// TwinCAT 3 PLC project Syn_Visu_Demo
// ProgramVersion: 3.1.4026.28
// libraries:
//   SynConfig,2.4.0.0,Syntegon Group
//   SynVisu,10.0.0.0,Syntegon Group
//   Tc3_Module,newest,Beckhoff Automation GmbH
//   Tc2_System, * (Beckhoff Automation GmbH)
// project tree:
//   / DEMO_GlobalConst.TcGVL, DEMO_GlobalVar.TcGVL, GVL_Config.TcGVL, GVL_Visu.TcGVL, TVisuDemo_Detection.TcDUT, TVisuDemo_Recipe.TcDUT
//   POUs/ PlcTask.TcTTO, P_VisuDemo.TcPOU, P_VisuDemoCartesian.TcPOU, P_VisuDemoCartesianAxes.TcPOU, P_VisuDemoDelta.TcPOU, P_VisuDemoFxx.TcPOU, P_VisuDemoIdh.TcPOU, P_VisuDemoMachine.TcPOU, P_VisuDemoSpacing.TcPOU, P_VisuDemoStress.TcPOU, _FC_DemoApproach.TcPOU
// (motion and I/O tree: see PLC project syn_visu)
// real-time tasks:
//   TASK PlcTask: cycle T#10ms, priority 20, ADS port 350
//   TASK TestTask: cycle T#10ms, priority 21, ADS port 351

CONFIGURATION Syn_Visu_Demo
    RESOURCE PLC ON TwinCAT3
        TASK PlcTask(INTERVAL := T#10ms, PRIORITY := 20);
        PROGRAM P_VisuDemo WITH PlcTask : P_VisuDemo;
    END_RESOURCE
END_CONFIGURATION

// ---- TVisuDemo_Detection.TcDUT
(* A raw detection as the demo's product generator makes it up and a vision system would report it: where the
   product lies (MCS), the belt position at that moment and its type. The demo's tracking latches it as Vision 1's. *)
TYPE TVisuDemo_Detection :
STRUCT
	Pose								: ST_VisuPlanarPose;	// MCS
	lr_BeltPosition						: LREAL;	// [mm] Infeed 1's belt position when it was seen
	udn_ProductType						: UDINT;	// [-]
END_STRUCT
END_TYPE

// ---- TVisuDemo_Recipe.TcDUT
(* The demo's effective recipe (ADR 0022): what P_VisuDemoMachine reads from its Syn_Config machine FB every cycle
   and the Delta application runs with: Infeed 1's belt, Delta 1 and the product generator before Vision 1. *)
TYPE TVisuDemo_Recipe :
STRUCT
	lr_BeltSpeed						: LREAL;	// [mm/s] Infeed 1
	lr_BeltAccel						: LREAL;	// [mm/s2] Infeed 1, also its deceleration
	lr_RobotSpeed						: LREAL;	// [%] Delta 1, of its maximum TCP speed
	lr_RobotAccel						: LREAL;	// [%] Delta 1, of its maximum TCP acceleration
	dn_PicksPerCycle					: DINT;	// [-] Delta 1 picks this many products before it places them: 1 or 2
	lr_Rate								: LREAL;	// [1/min] places the generator fills per minute at the recipe's belt speed
	dn_Lanes							: DINT;	// [-] pattern Lanes: lanes across the belt, 1..4; each product goes into one at random
	lr_LanePitch						: LREAL;	// [mm] between the lanes, centred on the belt
	dn_TypeMix							: DINT;	// [-] 0 = every type, 1 = boxes, 2 = round (can, oval)
	lr_ScatterX							: LREAL;	// [mm] at most along the belt, either way
	lr_ScatterY							: LREAL;	// [mm] at most across the belt, either way
	lr_ScatterRz						: LREAL;	// [deg] at most turned, either way
	lr_GapShare							: LREAL;	// [%] of the generator's places left empty
	dn_Seed								: DINT;	// [-] of the generator's pseudo-random numbers: the same seed gives the same products
	b_Feed								: BOOL;	// TRUE: the generator feeds products
	b_PatternLanes						: BOOL;	// TRUE: pattern Lanes (dn_Lanes, lr_LanePitch, unscattered); FALSE: Scattered (one lane, lr_Scatter*)
END_STRUCT
END_TYPE

// ---- DEMO_GlobalConst.TcGVL
(* Shared facts of the demo world: all applications use the same belt height and width, product and suction cup. *)
{attribute 'qualified_only'}
VAR_GLOBAL CONSTANT
	DEMO_lr_BELT_Z						: LREAL := 800;	// [mm] belt surface
	DEMO_lr_BELT_WIDTH					: LREAL := 400;	// [mm]
	DEMO_lr_PRODUCT_LENGTH				: LREAL := 120;	// [mm]
	DEMO_lr_PRODUCT_WIDTH				: LREAL := 80;	// [mm]
	DEMO_lr_PRODUCT_HEIGHT				: LREAL := 40;	// [mm]
	DEMO_lr_REMOVE_BEYOND_END			: LREAL := 300;	// [mm] register entries are dropped this far beyond the belt end
	(* Suction cup of Delta 1, the Fxx and IDH movers and the Cartesian robot: its grip point is where the products'
	   tops touch. *)
	DEMO_lr_CUP_DIAMETER				: LREAL := 40;	// [mm]
	DEMO_lr_CUP_HEIGHT					: LREAL := 50;	// [mm]
	(* Demo faults: every period one component or mover is in a fault for the duration. *)
	DEMO_lr_FAULT_PERIOD				: LREAL := 20;	// [s]
	DEMO_lr_FAULT_DURATION				: LREAL := 5;	// [s]
END_VAR

// ---- DEMO_GlobalVar.TcGVL
(* Shared runtime values of the demo. P_VisuDemo writes the cycle time and fault phase before it calls the
   applications; every application takes product ids from DEMO_udn_NextId. P_VisuDemoMachine, called first, writes
   the effective recipe, Infeed 1's belt speed and the reset; the Delta application reports a missed product. *)
{attribute 'qualified_only'}
VAR_GLOBAL
	DEMO_lr_Dt							: LREAL;	// [s] cycle time of the calling task
	DEMO_lr_FaultPhase					: LREAL;	// [s] 0..DEMO_lr_FAULT_PERIOD, drives the demo faults
	DEMO_udn_NextId						: UDINT := 1;	// [-] next product id, unique across all applications
	(* Load test (P_VisuDemoStress): products kept on the stress belt; 0 = off. Write it online. Once set, the stress
	   belt stays in the manifest until the next download or reset; set back to 0 it runs empty. *)
	DEMO_un_StressProducts				: UINT := 0;	// [-]
	(* Machine: the Delta application's sequence control (P_VisuDemoMachine, ADR 0022). *)
	DEMO_Recipe							: TVisuDemo_Recipe;	// the effective recipe
	DEMO_lr_Infeed1Speed				: LREAL;	// [mm/s] Infeed 1 now, ramped to the recipe's speed while running, to 0 when stopping
	DEMO_b_Reset						: BOOL;	// [-] one cycle: Reset accepted, Infeed 1 and Delta 1 start empty
	DEMO_b_Infeed1Missed				: BOOL;	// [-] a product passed Infeed 1's end unpicked a moment ago
END_VAR

// ---- GVL_Config.TcGVL
(* The application's config manifest (ADR 0017): the gateway finds the parameter FBs of Syn_Config at
   GVL_Config.stManifest. *)
{attribute 'qualified_only'}
VAR_GLOBAL
	stManifest : SynConfig.ST_ConfigManifest;
END_VAR

// ---- GVL_Visu.TcGVL
(* The application's manifest (ADR-0003): the gateway starts discovery at GVL_Visu.stManifest. Next to it the machine
   entry (protocol 22, ADR 0021): run state, simulation mode and machine messages, set by P_VisuDemo. *)
{attribute 'qualified_only'}
VAR_GLOBAL
	stManifest : ST_VisuManifest;
	stMachine : ST_VisuMachine;
END_VAR

// ---- POUs/P_VisuDemo.TcPOU
(****************************************************************************************************<br>
© Syntegon Group.<br>
All rights reserved, also regarding any disposal, exploitation, reproduction, editing, distribution,<br>
as well as in the event of applications for industrial property rights.<br>
*****************************************************************************************************<br>
DESCRIPTION:<br>
DEMO ONLY: independent sample applications side by side, for testing the gateway over ADS. All lines<br>
start at X = 0 and convey along +X. Each application is its own program:<br>
- P_VisuDemoDelta (Y = 0..1000): two infeeds, one outfeed, three Delta robots with different grippers; Infeed 1<br>
  is fed by a product generator and run, with Delta 1, by the sequence control P_VisuDemoMachine.<br>
- P_VisuDemoFxx (Y = 2500): an XTS loop above two belts evens out irregular gaps.<br>
- P_VisuDemoIdh (Y = 4100..4850): an XTS gantry picks in batches onto a tray belt.<br>
- P_VisuDemoCartesian (Y = 6500..7300): a Cartesian robot turns and tilts the products it places.<br>
- P_VisuDemoCartesianAxes (X = 4000, Y = 6500..7800): Cartesian robots without Y or without Z axis.<br>
- P_VisuDemoSpacing (Y = 9000): an XTS loop under one belt hands products back with a constant pitch.<br>
- P_VisuDemoStress (Y = 11000): load test with thousands of products, off unless DEMO_un_StressProducts is set.<br>
This program, called by PlcTask, sets the shared cycle time and fault phase (DEMO_GlobalVar), calls the machine's<br>
sequence control (recipe, commands, run state, machine messages: P_VisuDemoMachine) and then the applications.<br>
Part of the demo application Syn_Visu_Demo, which uses the Syn_Visu library like any machine project.<br>
****************************************************************************************************)
PROGRAM P_VisuDemo
VAR
	dn_TaskIndex						: DINT;
END_VAR

(****************************************************************************************************)
(* CYCLE TIME AND FAULT PHASE                                                                       *)
(****************************************************************************************************)
dn_TaskIndex := Tc2_System.GETCURTASKINDEXEX();
IF dn_TaskIndex > 0 THEN
	DEMO_GlobalVar.DEMO_lr_Dt := UDINT_TO_LREAL(TwinCAT_SystemInfoVarList._TaskInfo[dn_TaskIndex].CycleTime) * 1.0E-7;
ELSE
	DEMO_GlobalVar.DEMO_lr_Dt := 0.01;
END_IF
DEMO_GlobalVar.DEMO_lr_FaultPhase := DEMO_GlobalVar.DEMO_lr_FaultPhase + DEMO_GlobalVar.DEMO_lr_Dt;
IF DEMO_GlobalVar.DEMO_lr_FaultPhase >= DEMO_GlobalConst.DEMO_lr_FAULT_PERIOD THEN
	DEMO_GlobalVar.DEMO_lr_FaultPhase := DEMO_GlobalVar.DEMO_lr_FaultPhase - DEMO_GlobalConst.DEMO_lr_FAULT_PERIOD;
END_IF


(****************************************************************************************************)
(* MACHINE: recipe, commands and run state first, so the applications run with this cycle's values    *)
(****************************************************************************************************)
P_VisuDemoMachine();


(****************************************************************************************************)
(* APPLICATIONS                                                                                     *)
(****************************************************************************************************)
P_VisuDemoDelta();
P_VisuDemoFxx();
P_VisuDemoIdh();
P_VisuDemoCartesian();
P_VisuDemoCartesianAxes();
P_VisuDemoSpacing();
P_VisuDemoStress();

END_PROGRAM

// ---- POUs/P_VisuDemoMachine.TcPOU
(****************************************************************************************************<br>
© Syntegon Group.<br>
All rights reserved, also regarding any disposal, exploitation, reproduction, editing, distribution,<br>
as well as in the event of applications for industrial property rights.<br>
*****************************************************************************************************<br>
DESCRIPTION:<br>
DEMO ONLY: the minimal sequence control of the Delta application's Infeed 1 and Delta 1, as the Simulator drives it<br>
(ADR 0022). Its Syn_Config machine FB declares the recipe (Infeed 1's belt, Delta 1, the product pattern of the<br>
generator before Vision 1) and hands it Start, Stop and Reset; the effective recipe goes to DEMO_GlobalVar for<br>
P_VisuDemoDelta. Run states: STARTING ramps Infeed 1 up to the recipe's speed, RUNNING, STOPPING ramps it down,<br>
STOPPED; Delta 1 moves only as fast as its belt, so it halts with it. Start is accepted while stopped, Stop while<br>
starting or running, Reset while stopped: it empties Infeed 1 and Delta 1, restarts the generator from its seed and<br>
acknowledges the missed-product message and Delta 1's fault. The demo starts running and always reports simulation<br>
mode. It reports the machine to Syn_Visu (GVL_Visu.stMachine) with two machine messages: 'Reject bin almost full'<br>
about the reject unit for lr_REJECT_BIN_DURATION of every fault period, and 'Product missed' about Infeed 1. Its<br>
Syn_Config topology FB declares the demo's topology (ADR 0023, m_DeclareTopology). Called first by P_VisuDemo.<br>
****************************************************************************************************)
PROGRAM P_VisuDemoMachine
VAR
	fb_Machine							: _FB_VisuMachine;	// Syn_Visu: run state, simulation mode, machine messages
	fb_MachineParam						: SynConfig._FB_ConfigMachine;	// Syn_Config: recipe and commands
	fb_Topology							: SynConfig._FB_ConfigTopology;	// Syn_Config: the demo's topology (ADR 0023)
	e_RunState							: E_VisuRunState := E_VisuRunState.STARTING;	// the demo starts running
	lr_TargetSpeed						: LREAL;	// [mm/s] Infeed 1 ramps to this
	lr_RampStep							: LREAL;	// [mm/s] Infeed 1's speed change at most this cycle
END_VAR
VAR PERSISTENT
	RecipeSet							: SynConfig.ST_ConfigRecipeSet;	// the active recipe, kept over a restart
END_VAR
VAR CONSTANT
	(* Recipe fields, in the order they are declared: keep it, add new ones at the end. *)
	un_F_BELT_SPEED						: UINT := 1;
	un_F_BELT_ACCEL						: UINT := 2;
	un_F_ROBOT_SPEED					: UINT := 3;
	un_F_ROBOT_ACCEL					: UINT := 4;
	un_F_PICKS							: UINT := 5;
	un_F_RATE							: UINT := 6;
	un_F_LANES							: UINT := 7;
	un_F_LANE_PITCH						: UINT := 8;
	un_F_TYPE_MIX						: UINT := 9;
	un_F_SCATTER_X						: UINT := 10;
	un_F_SCATTER_Y						: UINT := 11;
	un_F_SCATTER_RZ						: UINT := 12;
	un_F_GAP_SHARE						: UINT := 13;
	un_F_SEED							: UINT := 14;
	un_F_FEED							: UINT := 15;
	un_F_PATTERN						: UINT := 16;
	(* Pattern: Scattered is 0, so a recipe saved before the field existed (its value 0) keeps the demo's old pattern. *)
	dn_PATTERN_SCATTERED				: DINT := 0;	// [-] Pattern: one lane, scattered
	dn_PATTERN_LANES					: DINT := 1;	// [-] Pattern: in lanes, unscattered
	udn_INFEED1_ID						: UDINT := 1;	// [-] manifest id of Infeed 1 (P_VisuDemoDelta)
	udn_DELTA1_ID						: UDINT := 10;	// [-] manifest id of Delta 1 (P_VisuDemoDelta)
	udn_REJECT_UNIT_ID					: UDINT := 60;	// [-] manifest id of the reject unit (P_VisuDemoDelta)
	udn_VISION1_ID						: UDINT := 50;	// [-] manifest id of Vision 1 (P_VisuDemoDelta)
	udn_MSG_REJECT_BIN					: UDINT := 1;	// [-] machine message: the reject bin is almost full
	udn_MSG_MISSED						: UDINT := 2;	// [-] machine message: a product passed Infeed 1 unpicked
	lr_REJECT_BIN_DURATION				: LREAL := 4;	// [s] the reject bin message is active from the start of every fault period
END_VAR

(****************************************************************************************************)
(* RECIPE (declaration idempotent, every cycle)                                                     *)
(****************************************************************************************************)
fb_MachineParam.m_Register(vio_Manifest := GVL_Config.stManifest, vi_udn_Id := 0);
m_DeclareFields();
(* The demo takes a recipe over at once; a machine would wait until it stands. *)
fb_MachineParam.m_Cycle(vio_Set := RecipeSet, vi_b_ApplyAllowed := TRUE);
DEMO_GlobalVar.DEMO_Recipe.lr_BeltSpeed := fb_MachineParam.m_Value(vi_un_Field := un_F_BELT_SPEED);
DEMO_GlobalVar.DEMO_Recipe.lr_BeltAccel := fb_MachineParam.m_Value(vi_un_Field := un_F_BELT_ACCEL);
DEMO_GlobalVar.DEMO_Recipe.lr_RobotSpeed := fb_MachineParam.m_Value(vi_un_Field := un_F_ROBOT_SPEED);
DEMO_GlobalVar.DEMO_Recipe.lr_RobotAccel := fb_MachineParam.m_Value(vi_un_Field := un_F_ROBOT_ACCEL);
DEMO_GlobalVar.DEMO_Recipe.dn_PicksPerCycle := fb_MachineParam.m_Integer(vi_un_Field := un_F_PICKS);
DEMO_GlobalVar.DEMO_Recipe.lr_Rate := fb_MachineParam.m_Value(vi_un_Field := un_F_RATE);
DEMO_GlobalVar.DEMO_Recipe.dn_Lanes := fb_MachineParam.m_Integer(vi_un_Field := un_F_LANES);
DEMO_GlobalVar.DEMO_Recipe.lr_LanePitch := fb_MachineParam.m_Value(vi_un_Field := un_F_LANE_PITCH);
DEMO_GlobalVar.DEMO_Recipe.dn_TypeMix := fb_MachineParam.m_Integer(vi_un_Field := un_F_TYPE_MIX);
DEMO_GlobalVar.DEMO_Recipe.lr_ScatterX := fb_MachineParam.m_Value(vi_un_Field := un_F_SCATTER_X);
DEMO_GlobalVar.DEMO_Recipe.lr_ScatterY := fb_MachineParam.m_Value(vi_un_Field := un_F_SCATTER_Y);
DEMO_GlobalVar.DEMO_Recipe.lr_ScatterRz := fb_MachineParam.m_Value(vi_un_Field := un_F_SCATTER_RZ);
DEMO_GlobalVar.DEMO_Recipe.lr_GapShare := fb_MachineParam.m_Value(vi_un_Field := un_F_GAP_SHARE);
DEMO_GlobalVar.DEMO_Recipe.dn_Seed := fb_MachineParam.m_Integer(vi_un_Field := un_F_SEED);
DEMO_GlobalVar.DEMO_Recipe.b_Feed := fb_MachineParam.m_Switch(vi_un_Field := un_F_FEED);
DEMO_GlobalVar.DEMO_Recipe.b_PatternLanes := fb_MachineParam.m_Integer(vi_un_Field := un_F_PATTERN) = dn_PATTERN_LANES;


(****************************************************************************************************)
(* TOPOLOGY (declaration and program values idempotent, every cycle)                                *)
(****************************************************************************************************)
fb_Topology.m_Register(vio_Manifest := GVL_Config.stManifest, vi_udn_Id := 0);
m_DeclareTopology();
fb_Topology.m_Cycle();


(****************************************************************************************************)
(* COMMANDS: the application decides                                                                *)
(****************************************************************************************************)
DEMO_GlobalVar.DEMO_b_Reset := FALSE;
CASE fb_MachineParam.m_Command() OF
	SynConfig.E_ConfigCommand.START:
		IF e_RunState = E_VisuRunState.STOPPED THEN
			e_RunState := E_VisuRunState.STARTING;
			fb_MachineParam.m_AnswerCommand(vi_b_Accepted := TRUE, vi_str_Reason := '');
		ELSE
			fb_MachineParam.m_AnswerCommand(vi_b_Accepted := FALSE, vi_str_Reason := 'The machine is not stopped');
		END_IF
	SynConfig.E_ConfigCommand.STOP:
		IF e_RunState = E_VisuRunState.STARTING OR e_RunState = E_VisuRunState.RUNNING THEN
			e_RunState := E_VisuRunState.STOPPING;
			fb_MachineParam.m_AnswerCommand(vi_b_Accepted := TRUE, vi_str_Reason := '');
		ELSE
			fb_MachineParam.m_AnswerCommand(vi_b_Accepted := FALSE, vi_str_Reason := 'The machine is not running');
		END_IF
	SynConfig.E_ConfigCommand.RESET:
		IF e_RunState = E_VisuRunState.STOPPED THEN
			DEMO_GlobalVar.DEMO_b_Reset := TRUE;
			fb_MachineParam.m_AnswerCommand(vi_b_Accepted := TRUE, vi_str_Reason := '');
		ELSE
			fb_MachineParam.m_AnswerCommand(vi_b_Accepted := FALSE, vi_str_Reason := 'Stop the machine first');
		END_IF
END_CASE


(****************************************************************************************************)
(* RUN STATE: Infeed 1 ramps up while starting and running, down while stopping                     *)
(****************************************************************************************************)
IF e_RunState = E_VisuRunState.STARTING OR e_RunState = E_VisuRunState.RUNNING THEN
	lr_TargetSpeed := DEMO_GlobalVar.DEMO_Recipe.lr_BeltSpeed;
ELSE
	lr_TargetSpeed := 0;
END_IF
lr_RampStep := DEMO_GlobalVar.DEMO_Recipe.lr_BeltAccel * DEMO_GlobalVar.DEMO_lr_Dt;
DEMO_GlobalVar.DEMO_lr_Infeed1Speed := _FC_DemoApproach(DEMO_GlobalVar.DEMO_lr_Infeed1Speed, lr_TargetSpeed, lr_RampStep);
IF e_RunState = E_VisuRunState.STARTING AND DEMO_GlobalVar.DEMO_lr_Infeed1Speed = lr_TargetSpeed THEN
	e_RunState := E_VisuRunState.RUNNING;
ELSIF e_RunState = E_VisuRunState.STOPPING AND DEMO_GlobalVar.DEMO_lr_Infeed1Speed = 0 THEN
	e_RunState := E_VisuRunState.STOPPED;
END_IF


(****************************************************************************************************)
(* REPORT: the machine to Syn_Visu                                                                  *)
(****************************************************************************************************)
fb_Machine.m_Register(vio_Machine := GVL_Visu.stMachine);
fb_Machine.m_SetRunState(vi_e_RunState := e_RunState, vi_str_Text := '');
fb_Machine.m_SetSimulation(vi_b_Simulation := TRUE);
fb_Machine.m_SetMessage(vi_udn_Id := udn_MSG_REJECT_BIN,
	vi_b_Active := DEMO_GlobalVar.DEMO_lr_FaultPhase < lr_REJECT_BIN_DURATION, vi_e_Severity := E_VisuMessageSeverity.WARNING,
	vi_str_Text := 'Reject bin almost full', vi_udn_ComponentId := udn_REJECT_UNIT_ID);
fb_Machine.m_SetMessage(vi_udn_Id := udn_MSG_MISSED, vi_b_Active := DEMO_GlobalVar.DEMO_b_Infeed1Missed,
	vi_e_Severity := E_VisuMessageSeverity.WARNING, vi_str_Text := 'Product missed', vi_udn_ComponentId := udn_INFEED1_ID);

(****************************************************************************************************<br>
© Syntegon Group.<br>
All rights reserved, also regarding any disposal, exploitation, reproduction, editing, distribution,<br>
as well as in the event of applications for industrial property rights.<br>
*****************************************************************************************************<br>
DESCRIPTION:<br>
The demo's recipe fields: Infeed 1's belt, Delta 1 and the product pattern of the generator before Vision 1 (for<br>
the whole machine), each with a description and some with a label of their own (Syn_Config 2.2.0). The pattern is<br>
Lanes or Scattered: the lane fields apply only to Lanes, the scatter fields only to Scattered, so the Simulator<br>
shows only the fields of the chosen one. The program values give the pattern the demo had before its recipe: one<br>
lane, 60 products a minute at 150 mm/s, every product type, scattered across the belt and turned. Rate counts the<br>
generator's places a minute at the recipe's belt speed: the pattern keeps its spacing while the belt ramps.<br>
****************************************************************************************************)
METHOD PRIVATE m_DeclareFields
fb_MachineParam.m_DeclareField(vi_un_Field := un_F_BELT_SPEED, vi_str_Name := 'BeltSpeed', vi_udn_Group := udn_INFEED1_ID,
	vi_e_Type := SynConfig.E_ConfigFieldType.NUMBER, vi_str_Unit := 'mm/s', vi_lr_Min := 10, vi_lr_Max := 500,
	vi_lr_ProgramValue := 150);
fb_MachineParam.m_DeclareField(vi_un_Field := un_F_BELT_ACCEL, vi_str_Name := 'BeltAcceleration', vi_udn_Group := udn_INFEED1_ID,
	vi_e_Type := SynConfig.E_ConfigFieldType.NUMBER, vi_str_Unit := 'mm/s2', vi_lr_Min := 50, vi_lr_Max := 2000,
	vi_lr_ProgramValue := 300);
fb_MachineParam.m_DeclareField(vi_un_Field := un_F_ROBOT_SPEED, vi_str_Name := 'RobotSpeed', vi_udn_Group := udn_DELTA1_ID,
	vi_e_Type := SynConfig.E_ConfigFieldType.NUMBER, vi_str_Unit := '%', vi_lr_Min := 10, vi_lr_Max := 100,
	vi_lr_ProgramValue := 100);
fb_MachineParam.m_DeclareField(vi_un_Field := un_F_ROBOT_ACCEL, vi_str_Name := 'RobotAcceleration', vi_udn_Group := udn_DELTA1_ID,
	vi_e_Type := SynConfig.E_ConfigFieldType.NUMBER, vi_str_Unit := '%', vi_lr_Min := 10, vi_lr_Max := 100,
	vi_lr_ProgramValue := 100);
fb_MachineParam.m_DeclareField(vi_un_Field := un_F_PICKS, vi_str_Name := 'PicksPerCycle', vi_udn_Group := udn_DELTA1_ID,
	vi_e_Type := SynConfig.E_ConfigFieldType.INTEGER, vi_str_Unit := '', vi_lr_Min := 1, vi_lr_Max := 2,
	vi_lr_ProgramValue := 2);
fb_MachineParam.m_DeclareField(vi_un_Field := un_F_RATE, vi_str_Name := 'Rate', vi_udn_Group := 0,
	vi_e_Type := SynConfig.E_ConfigFieldType.NUMBER, vi_str_Unit := '1/min', vi_lr_Min := 1, vi_lr_Max := 120,
	vi_lr_ProgramValue := 60);
fb_MachineParam.m_DeclareField(vi_un_Field := un_F_LANES, vi_str_Name := 'Lanes', vi_udn_Group := 0,
	vi_e_Type := SynConfig.E_ConfigFieldType.INTEGER, vi_str_Unit := '', vi_lr_Min := 1, vi_lr_Max := 4,
	vi_lr_ProgramValue := 1);
fb_MachineParam.m_DeclareField(vi_un_Field := un_F_LANE_PITCH, vi_str_Name := 'LanePitch', vi_udn_Group := 0,
	vi_e_Type := SynConfig.E_ConfigFieldType.NUMBER, vi_str_Unit := 'mm', vi_lr_Min := 0, vi_lr_Max := 150,
	vi_lr_ProgramValue := 90);
fb_MachineParam.m_DeclareField(vi_un_Field := un_F_TYPE_MIX, vi_str_Name := 'TypeMix', vi_udn_Group := 0,
	vi_e_Type := SynConfig.E_ConfigFieldType.CHOICE, vi_str_Unit := '', vi_lr_Min := 0, vi_lr_Max := 0,
	vi_lr_ProgramValue := 0);
fb_MachineParam.m_SetChoice(vi_un_Field := un_F_TYPE_MIX, vi_un_Value := 0, vi_str_Text := 'Every type');
fb_MachineParam.m_SetChoice(vi_un_Field := un_F_TYPE_MIX, vi_un_Value := 1, vi_str_Text := 'Boxes');
fb_MachineParam.m_SetChoice(vi_un_Field := un_F_TYPE_MIX, vi_un_Value := 2, vi_str_Text := 'Round');
fb_MachineParam.m_DeclareField(vi_un_Field := un_F_SCATTER_X, vi_str_Name := 'ScatterX', vi_udn_Group := 0,
	vi_e_Type := SynConfig.E_ConfigFieldType.NUMBER, vi_str_Unit := 'mm', vi_lr_Min := 0, vi_lr_Max := 50,
	vi_lr_ProgramValue := 0);
fb_MachineParam.m_DeclareField(vi_un_Field := un_F_SCATTER_Y, vi_str_Name := 'ScatterY', vi_udn_Group := 0,
	vi_e_Type := SynConfig.E_ConfigFieldType.NUMBER, vi_str_Unit := 'mm', vi_lr_Min := 0, vi_lr_Max := 100,
	vi_lr_ProgramValue := 80);
fb_MachineParam.m_DeclareField(vi_un_Field := un_F_SCATTER_RZ, vi_str_Name := 'ScatterRz', vi_udn_Group := 0,
	vi_e_Type := SynConfig.E_ConfigFieldType.NUMBER, vi_str_Unit := 'deg', vi_lr_Min := 0, vi_lr_Max := 90,
	vi_lr_ProgramValue := 30);
fb_MachineParam.m_DeclareField(vi_un_Field := un_F_GAP_SHARE, vi_str_Name := 'GapShare', vi_udn_Group := 0,
	vi_e_Type := SynConfig.E_ConfigFieldType.NUMBER, vi_str_Unit := '%', vi_lr_Min := 0, vi_lr_Max := 90,
	vi_lr_ProgramValue := 0);
fb_MachineParam.m_DeclareField(vi_un_Field := un_F_SEED, vi_str_Name := 'Seed', vi_udn_Group := 0,
	vi_e_Type := SynConfig.E_ConfigFieldType.INTEGER, vi_str_Unit := '', vi_lr_Min := 1, vi_lr_Max := 999999,
	vi_lr_ProgramValue := 12345);
fb_MachineParam.m_DeclareField(vi_un_Field := un_F_FEED, vi_str_Name := 'Feed', vi_udn_Group := 0,
	vi_e_Type := SynConfig.E_ConfigFieldType.SWITCH, vi_str_Unit := '', vi_lr_Min := 0, vi_lr_Max := 0,
	vi_lr_ProgramValue := 1);
fb_MachineParam.m_DeclareField(vi_un_Field := un_F_PATTERN, vi_str_Name := 'Pattern', vi_udn_Group := 0,
	vi_e_Type := SynConfig.E_ConfigFieldType.CHOICE, vi_str_Unit := '', vi_lr_Min := 0, vi_lr_Max := 0,
	vi_lr_ProgramValue := DINT_TO_LREAL(dn_PATTERN_SCATTERED));
fb_MachineParam.m_SetChoice(vi_un_Field := un_F_PATTERN, vi_un_Value := DINT_TO_UINT(dn_PATTERN_SCATTERED), vi_str_Text := 'Scattered');
fb_MachineParam.m_SetChoice(vi_un_Field := un_F_PATTERN, vi_un_Value := DINT_TO_UINT(dn_PATTERN_LANES), vi_str_Text := 'Lanes');


(****************************************************************************************************)
(* TEXTS: label ('' = the name put into words) and description                                     *)
(****************************************************************************************************)
fb_MachineParam.m_SetText(vi_un_Field := un_F_BELT_SPEED, vi_str_Label := '',
	vi_str_Description := 'Speed Infeed 1 ramps up to while the machine runs');
fb_MachineParam.m_SetText(vi_un_Field := un_F_BELT_ACCEL, vi_str_Label := '',
	vi_str_Description := 'How fast Infeed 1 speeds up after Start and slows down after Stop');
fb_MachineParam.m_SetText(vi_un_Field := un_F_ROBOT_SPEED, vi_str_Label := '',
	vi_str_Description := 'Delta 1 moves at this share of its maximum TCP speed');
fb_MachineParam.m_SetText(vi_un_Field := un_F_ROBOT_ACCEL, vi_str_Label := '',
	vi_str_Description := 'Delta 1 accelerates at this share of its maximum TCP acceleration');
fb_MachineParam.m_SetText(vi_un_Field := un_F_PICKS, vi_str_Label := '',
	vi_str_Description := 'Products Delta 1 picks before it places them');
fb_MachineParam.m_SetText(vi_un_Field := un_F_RATE, vi_str_Label := '',
	vi_str_Description := 'Places the generator fills a minute at the belt speed of the recipe');
fb_MachineParam.m_SetText(vi_un_Field := un_F_PATTERN, vi_str_Label := '',
	vi_str_Description := 'Scattered: one lane, scattered along, across and turned. Lanes: in lanes, unscattered');
fb_MachineParam.m_SetText(vi_un_Field := un_F_LANES, vi_str_Label := '',
	vi_str_Description := 'Lanes across the belt; each product goes into one at random');
fb_MachineParam.m_SetText(vi_un_Field := un_F_LANE_PITCH, vi_str_Label := '',
	vi_str_Description := 'Distance between the lanes, centred on the belt');
fb_MachineParam.m_SetText(vi_un_Field := un_F_TYPE_MIX, vi_str_Label := '',
	vi_str_Description := 'Which product types the generator feeds');
fb_MachineParam.m_SetText(vi_un_Field := un_F_SCATTER_X, vi_str_Label := 'Scatter along',
	vi_str_Description := 'A product lies at most this far before or behind its place');
fb_MachineParam.m_SetText(vi_un_Field := un_F_SCATTER_Y, vi_str_Label := 'Scatter across',
	vi_str_Description := 'A product lies at most this far beside the middle of the belt');
fb_MachineParam.m_SetText(vi_un_Field := un_F_SCATTER_RZ, vi_str_Label := 'Scatter turn',
	vi_str_Description := 'A product is turned at most this far either way');
fb_MachineParam.m_SetText(vi_un_Field := un_F_GAP_SHARE, vi_str_Label := 'Gaps',
	vi_str_Description := 'Share of the places left empty');
fb_MachineParam.m_SetText(vi_un_Field := un_F_SEED, vi_str_Label := 'Random seed',
	vi_str_Description := 'The same seed gives the same products; a new one starts the pattern again');
fb_MachineParam.m_SetText(vi_un_Field := un_F_FEED, vi_str_Label := '',
	vi_str_Description := 'Off: the generator feeds no products');


(****************************************************************************************************)
(* CONDITIONS: the lane fields only for Lanes, the scatter fields only for Scattered                *)
(****************************************************************************************************)
fb_MachineParam.m_SetVisibleWhen(vi_un_Field := un_F_LANES, vi_un_OnField := un_F_PATTERN, vi_dn_Value := dn_PATTERN_LANES);
fb_MachineParam.m_SetVisibleWhen(vi_un_Field := un_F_LANE_PITCH, vi_un_OnField := un_F_PATTERN, vi_dn_Value := dn_PATTERN_LANES);
fb_MachineParam.m_SetVisibleWhen(vi_un_Field := un_F_SCATTER_X, vi_un_OnField := un_F_PATTERN, vi_dn_Value := dn_PATTERN_SCATTERED);
fb_MachineParam.m_SetVisibleWhen(vi_un_Field := un_F_SCATTER_Y, vi_un_OnField := un_F_PATTERN, vi_dn_Value := dn_PATTERN_SCATTERED);
fb_MachineParam.m_SetVisibleWhen(vi_un_Field := un_F_SCATTER_RZ, vi_un_OnField := un_F_PATTERN, vi_dn_Value := dn_PATTERN_SCATTERED);
END_METHOD

(****************************************************************************************************<br>
© Syntegon Group.<br>
All rights reserved, also regarding any disposal, exploitation, reproduction, editing, distribution,<br>
as well as in the event of applications for industrial property rights.<br>
*****************************************************************************************************<br>
DESCRIPTION:<br>
DEMO ONLY: the demo's topology (ADR 0023) in the words of the RPP application. The line TCAT1 (root) holds the cell<br>
MPS1, which holds the transport TBL1 (Infeed 1), the pick-and-place handling PPH1 (Delta 1) taking its products<br>
from TBL1 and the vision unit DET1 (Vision 1) looking at TBL1. PPH2 belongs to the full build-out but has no<br>
parent: it is not in use. Idempotent, every cycle.<br>
****************************************************************************************************)
METHOD PRIVATE m_DeclareTopology
VAR CONSTANT
	un_K_LINE							: UINT := 1;	// [-] kinds
	un_K_CELL							: UINT := 2;
	un_K_TRANSPORT						: UINT := 3;
	un_K_PPH							: UINT := 4;
	un_K_DET							: UINT := 5;
	un_R_INFEED1						: UINT := 1;	// [-] roles
	un_R_TRANSPORT						: UINT := 2;
	dn_TCAT1							: DINT := 1;	// [-] nodes, numbered like the RPP application's contexts
	dn_MPS1								: DINT := 10;
	dn_PPH1								: DINT := 21;
	dn_PPH2								: DINT := 22;
	dn_TBL1								: DINT := 30;
	dn_DET1								: DINT := 60;
END_VAR
fb_Topology.m_DeclareKind(vi_un_Kind := un_K_LINE, vi_str_Name := 'Line');
fb_Topology.m_DeclareKind(vi_un_Kind := un_K_CELL, vi_str_Name := 'Cell');
fb_Topology.m_DeclareKind(vi_un_Kind := un_K_TRANSPORT, vi_str_Name := 'Transport');
fb_Topology.m_DeclareKind(vi_un_Kind := un_K_PPH, vi_str_Name := 'PPH');
fb_Topology.m_DeclareKind(vi_un_Kind := un_K_DET, vi_str_Name := 'DET');
fb_Topology.m_AllowParent(vi_un_Kind := un_K_CELL, vi_un_ParentKind := un_K_LINE);
fb_Topology.m_AllowParent(vi_un_Kind := un_K_TRANSPORT, vi_un_ParentKind := un_K_CELL);
fb_Topology.m_AllowParent(vi_un_Kind := un_K_PPH, vi_un_ParentKind := un_K_CELL);
fb_Topology.m_AllowParent(vi_un_Kind := un_K_DET, vi_un_ParentKind := un_K_CELL);
fb_Topology.m_DeclareRole(vi_un_Role := un_R_INFEED1, vi_str_Name := 'Infeed1', vi_un_HolderKind := un_K_PPH, vi_b_Required := TRUE);
fb_Topology.m_AllowTarget(vi_un_Role := un_R_INFEED1, vi_un_TargetKind := un_K_TRANSPORT);
fb_Topology.m_DeclareRole(vi_un_Role := un_R_TRANSPORT, vi_str_Name := 'Transport', vi_un_HolderKind := un_K_DET, vi_b_Required := TRUE);
fb_Topology.m_AllowTarget(vi_un_Role := un_R_TRANSPORT, vi_un_TargetKind := un_K_TRANSPORT);

fb_Topology.m_DeclareNode(vi_dn_Id := dn_TCAT1, vi_str_Name := 'TCAT1', vi_un_Kind := un_K_LINE);
fb_Topology.m_DeclareNode(vi_dn_Id := dn_MPS1, vi_str_Name := 'MPS1', vi_un_Kind := un_K_CELL);
fb_Topology.m_DeclareNode(vi_dn_Id := dn_TBL1, vi_str_Name := 'TBL1', vi_un_Kind := un_K_TRANSPORT);
fb_Topology.m_DeclareNode(vi_dn_Id := dn_PPH1, vi_str_Name := 'PPH1', vi_un_Kind := un_K_PPH);
fb_Topology.m_DeclareNode(vi_dn_Id := dn_PPH2, vi_str_Name := 'PPH2', vi_un_Kind := un_K_PPH);
fb_Topology.m_DeclareNode(vi_dn_Id := dn_DET1, vi_str_Name := 'DET1', vi_un_Kind := un_K_DET);
fb_Topology.m_AddComponent(vi_dn_Node := dn_TBL1, vi_udn_ComponentId := udn_INFEED1_ID);
fb_Topology.m_AddComponent(vi_dn_Node := dn_PPH1, vi_udn_ComponentId := udn_DELTA1_ID);
fb_Topology.m_AddComponent(vi_dn_Node := dn_DET1, vi_udn_ComponentId := udn_VISION1_ID);
fb_Topology.m_SetRoot(vi_dn_Node := dn_TCAT1);

(* Program values: the links the demo runs with. *)
fb_Topology.m_SetParent(vi_dn_Node := dn_MPS1, vi_dn_Parent := dn_TCAT1);
fb_Topology.m_SetParent(vi_dn_Node := dn_TBL1, vi_dn_Parent := dn_MPS1);
fb_Topology.m_SetParent(vi_dn_Node := dn_PPH1, vi_dn_Parent := dn_MPS1);
fb_Topology.m_SetParent(vi_dn_Node := dn_DET1, vi_dn_Parent := dn_MPS1);
fb_Topology.m_Link(vi_dn_Node := dn_PPH1, vi_un_Role := un_R_INFEED1, vi_dn_Target := dn_TBL1);
fb_Topology.m_Link(vi_dn_Node := dn_DET1, vi_un_Role := un_R_TRANSPORT, vi_dn_Target := dn_TBL1);
END_METHOD

END_PROGRAM

// ---- POUs/_FC_DemoApproach.TcPOU
(****************************************************************************************************<br>
© Syntegon Group.<br>
All rights reserved, also regarding any disposal, exploitation, reproduction, editing, distribution,<br>
as well as in the event of applications for industrial property rights.<br>
*****************************************************************************************************<br>
DESCRIPTION:<br>
Moves vi_lr_Value towards vi_lr_Goal by at most vi_lr_Step. Lands exactly on the goal, so callers may compare<br>
the result with the goal for equality.<br>
****************************************************************************************************)
FUNCTION _FC_DemoApproach : LREAL
VAR_INPUT
	vi_lr_Value							: LREAL;
	vi_lr_Goal							: LREAL;
	vi_lr_Step							: LREAL;	// >= 0
END_VAR

IF ABS(vi_lr_Goal - vi_lr_Value) <= vi_lr_Step THEN
	_FC_DemoApproach := vi_lr_Goal;
ELSIF vi_lr_Goal > vi_lr_Value THEN
	_FC_DemoApproach := vi_lr_Value + vi_lr_Step;
ELSE
	_FC_DemoApproach := vi_lr_Value - vi_lr_Step;
END_IF

END_FUNCTION

// ---- POUs/P_VisuDemoDelta.TcPOU
(****************************************************************************************************<br>
© Syntegon Group.<br>
All rights reserved, also regarding any disposal, exploitation, reproduction, editing, distribution,<br>
as well as in the event of applications for industrial property rights.<br>
*****************************************************************************************************<br>
DESCRIPTION:<br>
DEMO ONLY: Delta application (Y = 0..1000). Two infeed conveyors (Y = 0 and Y = 1000) and an outfeed between<br>
them (Y = 500), three Delta robots one after another (X = 1500, 2500, 3500) picking from the infeeds and placing<br>
onto the outfeed. Some products are deliberately missed. Each Delta has a different gripper:<br>
- Delta 1: two suction cups beside the flange that turn about Rz; it picks two products and places both at once.<br>
- Delta 2: one finger that turns about Rz and tilts about Rx while carrying.<br>
- Delta 3: five fingers around the flange that close when picking and open when placing.<br>
Products come in five types of different size and shape (boxes, a can, an oval, a pouch), mixed on both infeeds;<br>
Delta 1 picks a pair of one type, Delta 3 closes its fingers around the product's outline. A product put down<br>
on the outfeed leaves the infeed's register.<br>
A vision system over infeed 1 detects its products in the middle of its field of view and marks every tenth as a<br>
sample (product mark 1, 'Sample'), which stays marked on the outfeed; a light barrier on<br>
infeed 2 detects them at their front edge, its beam lighting up while a product interrupts it.<br>
A reject unit (station) at the outfeed rejects every fifth product passing it: its pusher lights up and the<br>
product is off the belt shortly after.<br>
Delta 1 is in a fault now and then.<br>
Infeed 1 and Delta 1 run under the sequence control P_VisuDemoMachine (ADR 0022): Infeed 1 at its ramped speed, its<br>
products from the product generator (m_Generate: the recipe's pattern, deterministic from its seed) latched as<br>
Vision 1's (m_Track); Delta 1 as fast as its belt and recipe allow (m_Delta1Step), picking as many products per<br>
cycle as the recipe says. Reset (m_Reset) empties Infeed 1 and Delta 1 and acknowledges Delta 1's fault; a product<br>
passing Infeed 1 unpicked raises 'Product missed' (m_Missed). Called by P_VisuDemo.<br>
****************************************************************************************************)
PROGRAM P_VisuDemoDelta
VAR
	fb_Infeed1							: _FB_VisuConveyor;
	fb_Infeed2							: _FB_VisuConveyor;
	fb_Outfeed							: _FB_VisuConveyor;
	fb_Delta1							: _FB_VisuDelta;
	fb_Delta2							: _FB_VisuDelta;
	fb_Delta3							: _FB_VisuDelta;
	fb_Vision1							: _FB_VisuVision;	// over infeed 1
	fb_Barrier2							: _FB_VisuSensor;	// light barrier on infeed 2
	fb_RejectUnit						: _FB_VisuStation;	// at the outfeed

	(* Syn_Config (ADR 0017): Infeed 1, Delta 1 and Vision 1 run with the parameter sets the configurator writes,
	   else with their program values. The demo allows taking a set over at once; a machine would wait until it
	   stands. *)
	fb_Infeed1Param						: SynConfig._FB_ConfigConveyor;
	fb_Delta1Param						: SynConfig._FB_ConfigDelta;
	fb_Vision1Param						: SynConfig._FB_ConfigVision;
	Infeed1Default						: SynConfig.ST_ConfigConveyorParam;	// program values of Infeed 1
	Vision1Default						: SynConfig.ST_ConfigBodyComponentParam;	// program values of Vision 1
	RobotDefault						: SynConfig.ST_ConfigDeltaParam;	// program values of the Delta being configured
	Zone								: ST_VisuZone;	// Delta 1's pick zone on infeed 1, from its parameter set
	lr_AllocStart						: LREAL;	// [mm] MCS X where the current robot's allocation area on the current infeed starts
	lr_AllocEnd							: LREAL;	// [mm] MCS X where it ends
	n_Zone								: INT;

	(* Reject unit *)
	un_RejectPassed						: UINT;	// [-] products that passed the reject unit
	udn_RejectPushing					: UDINT;	// [-] product being pushed off, 0 = none
	lr_RejectLeft						: LREAL;	// [s] until the product being pushed is off the belt

	(* Conveyors *)
	lr_Dt								: LREAL;	// [s] cycle time
	udn_Seed							: UDINT := 12345;	// [-] pseudo random generator state
	lr_BeltPosition						: ARRAY[0..2] OF LREAL;	// [mm] infeed 1, infeed 2, outfeed
	lr_SinceSpawn2						: LREAL := 0.3;	// [s] since the last product on infeed 2
	un_Vision1Latches					: UINT;	// [-] products Vision 1 latched: every un_SAMPLE_EVERY-th is a sample
	fb_RefBelt							: REFERENCE TO _FB_VisuConveyor;
	BeltPose							: ST_VisuPose;
	LatchPose							: ST_VisuPlanarPose;
	n_Belt								: INT;
	lr_Random							: LREAL;	// [-] 0..1
	udn_Type							: UDINT;	// [-] product type, 1..udn_TYPE_COUNT
	DetectorPose						: ST_VisuPose;	// lens of the vision system, head of the light barrier
	b_BeamInterrupted					: BOOL;	// a product on infeed 2 covers the light barrier's beam

	(* Per Delta robot *)
	n_Phase								: ARRAY[0..2] OF INT;
	udn_TargetId						: ARRAY[0..2] OF UDINT;	// [-] product being approached, 0 = none
	n_TargetBelt						: ARRAY[0..2] OF INT;	// [-] 0 = infeed 1, 1 = infeed 2
	Tcp									: ARRAY[0..2] OF ST_VisuPosition;	// the gripper flange
	b_TcpInitialised					: ARRAY[0..2] OF BOOL;
	lr_ToolRz							: ARRAY[0..2] OF LREAL;	// [deg] tool rotation about MCS Z (4th axis)
	udn_Held							: ARRAY[0..2, 0..1] OF UDINT;	// [-] carried product ids per slot (Delta 1 carries two)
	n_HeldBelt							: ARRAY[0..2, 0..1] OF INT;	// [-] infeed of each carried product: 0 = infeed 1, 1 = infeed 2
	udn_HeldType						: ARRAY[0..2, 0..1] OF UDINT;	// [-] product type of each carried product
	un_HeldMark							: ARRAY[0..2, 0..1] OF UINT;	// [-] product mark of each carried product, 0 = none
	lr_HeldHeight						: LREAL;	// [mm] height of the product carried or approached
	n_HeldCount							: ARRAY[0..2] OF INT;
	lr_TiltRx							: LREAL;	// [deg] Delta 2: finger tilt about its X
	lr_Spread							: LREAL := 130;	// [mm] Delta 3: finger distance from the flange
	lr_SpreadClosed						: LREAL := 82;	// [mm] Delta 3: finger distance closed around the current product
	n_Finger							: INT;	// [-] finger used for the current pick, 0 = the flange
	n_FingerCount						: INT;
	n_Slot								: INT;
	lr_GripHeight						: LREAL;	// [mm] flange above the grip point of the finger used
	Grip								: ST_VisuPosition;	// MCS offset flange -> grip point of the finger used
	fb_RefRobot							: REFERENCE TO _FB_VisuDelta;
	BasePose							: ST_VisuPose;
	Product								: ST_VisuProduct;
	ProductPose							: ST_VisuPlanarPose;
	SetpointTcp							: ST_VisuPosition;
	b_Found								: BOOL;
	n_Robot								: INT;
	un_Index							: UINT;
	lr_BaseX							: LREAL;	// [mm]
	lr_Step								: LREAL;	// [mm] TCP travel per cycle
	lr_X								: LREAL;	// [mm] target
	lr_Y								: LREAL;	// [mm] target
	lr_TopZ								: LREAL;	// [mm] top of the target product
	lr_TargetRz							: LREAL;	// [deg]
	un_Placed							: ARRAY[0..2] OF UINT;	// [-] times each robot has put its products down
	lr_PlaceWait						: ARRAY[0..2] OF LREAL;	// [s] waited above the place position
	b_FarPlace							: BOOL;	// the current robot places far downstream this time

	(* Sequence control (P_VisuDemoMachine, recipe): Infeed 1 at its ramped speed, Delta 1 as fast as its belt and its
	   recipe allow, the product generator before Vision 1. *)
	lr_Delta1Speed						: LREAL;	// [mm/s] Delta 1's TCP speed now, ramped
	udn_GenRandom						: UDINT;	// [-] the generator's pseudo-random numbers, started from the recipe's seed
	dn_GenSeed							: DINT;	// [-] the seed they started from; another seed or a reset starts them again
	lr_GenTravel						: LREAL;	// [mm] Infeed 1's travel since the generator's last place
	lr_MissedLeft						: LREAL;	// [s] the missed-product message stays this long
	Detection							: TVisuDemo_Detection;	// the generator's detection this cycle, latched by m_Track
	b_FaultAcknowledged					: BOOL;	// [-] Reset acknowledged Delta 1's fault until the next fault period
END_VAR
VAR PERSISTENT
	Infeed1Set							: SynConfig.ST_ConfigConveyorSet;	// active parameter set of Infeed 1, kept over a restart
	Delta1Set							: SynConfig.ST_ConfigDeltaSet;	// active parameter set of Delta 1
	Vision1Set							: SynConfig.ST_ConfigBodyComponentSet;	// active parameter set of Vision 1
END_VAR
VAR CONSTANT
	lr_BELT_LENGTH						: LREAL := 5000;	// [mm]
	lr_INFEED_SPEED						: LREAL := 150;	// [mm/s]
	lr_OUTFEED_SPEED					: LREAL := 300;	// [mm/s] two infeeds' products, 150 mm apart
	lr_SPAWN_INTERVAL					: LREAL := 1.0;	// [s] per infeed: 150 mm apart, the longest product type
	(* Product types, the same on every belt; type 1 is the standard product of the other demo applications. *)
	(* 1, 2: boxes; 3: a round can; 4: an oval; 5: a pouch with rounded edges. *)
	udn_TYPE_COUNT						: UDINT := 5;
	e_TYPE_SHAPE						: ARRAY[1..5] OF E_VisuProductShape := [E_VisuProductShape.BOX, E_VisuProductShape.BOX,
											E_VisuProductShape.CYLINDER, E_VisuProductShape.CYLINDER,
											E_VisuProductShape.ROUNDED_BOX];
	lr_TYPE_LENGTH						: ARRAY[1..5] OF LREAL := [120, 150, 90, 110, 140];	// [mm] along the conveying direction (a cylinder: diameter)
	lr_TYPE_WIDTH						: ARRAY[1..5] OF LREAL := [80, 100, 90, 70, 90];	// [mm] across (a cylinder: diameter)
	lr_TYPE_HEIGHT						: ARRAY[1..5] OF LREAL := [40, 45, 60, 45, 40];	// [mm] at least lr_RING_HEIGHT
	lr_TYPE_CORNER_RADIUS				: ARRAY[1..5] OF LREAL := [0, 0, 0, 0, 20];	// [mm] rounded edges of a rounded box
	lr_INFEED1_Y						: LREAL := 0;	// [mm]
	lr_INFEED2_Y						: LREAL := 1000;	// [mm]
	lr_OUTFEED_Y						: LREAL := 500;	// [mm]
	(* Each belt's coordinate system: infeed 1 at its start, infeed 2 at its end, the outfeed under Delta 1.
	   Zones on a belt are given from its origin. *)
	lr_INFEED2_ORIGIN_X					: LREAL := 5000;	// [mm] from the belt start
	lr_OUTFEED_ORIGIN_X					: LREAL := 1500;	// [mm] from the belt start
	(* Detectors *)
	lr_VISION_X							: LREAL := 300;	// [mm] lens over infeed 1, middle of the field of view
	lr_VISION_FIELD						: LREAL := 400;	// [mm] field of view on the belt, along and across
	lr_VISION_DISTANCE					: LREAL := 800;	// [mm] lens above the belt
	lr_BARRIER_X						: LREAL := 300;	// [mm] beam across infeed 2
	lr_BARRIER_HEIGHT					: LREAL := 20;	// [mm] beam above the belt
	lr_BARRIER_BEAM						: LREAL := 500;	// [mm] from the head at the belt edge across the belt
	un_SAMPLE_EVERY						: UINT := 10;	// [-] Vision 1 marks every n-th product as a sample
	un_SAMPLE_MARK						: UINT := 1;	// [-] product mark of a sample, named 'Sample'
	(* Reject unit, behind the last robot *)
	lr_REJECT_X							: LREAL := 4500;	// [mm] MCS X of its pusher
	un_REJECT_EVERY						: UINT := 5;	// [-] every n-th product is rejected
	lr_REJECT_PUSH_TIME					: LREAL := 0.3;	// [s] the pusher pushes a product off the belt
	lr_ROBOT1_X							: LREAL := 1500;	// [mm]
	lr_ROBOT_PITCH						: LREAL := 1000;	// [mm] distance between robots along X
	lr_ROBOT_Y							: LREAL := 500;	// [mm]
	lr_ROBOT_Z							: LREAL := 1900;	// [mm]
	lr_TCP_SPEED						: LREAL := 2500;	// [mm/s]
	lr_HOVER							: LREAL := 120;	// [mm]
	lr_PICK_HALF_ZONE					: LREAL := 400;	// [mm]
	lr_PICK_HALF_LANE					: LREAL := 130;	// [mm] pick zones only cover the lane the products come in on
	lr_PLACE_HALF_ZONE					: LREAL := 300;	// [mm]
	lr_ALLOCATION_OFFSET				: LREAL := 300;	// [mm] products are allocated only up to this distance before the pick zone end
	lr_LEAD								: LREAL := 7.5;	// [mm] the robot leads the moving product
	(* Demo limit violation: Delta 2 puts every sixth time down far downstream and waits there for a gap on the
	   outfeed. Its TCP limit area then reaches into Delta 3's limit area and out of its own. *)
	un_FAR_PLACE_EVERY					: UINT := 6;	// [-]
	lr_FAR_PLACE_OFFSET					: LREAL := 480;	// [mm] downstream of its base
	lr_FAR_PLACE_WAIT					: LREAL := 0.8;	// [s]
	lr_FAULT_START						: LREAL := 4;	// [s] start of the Delta 1 fault in the fault period
	(* Grippers *)
	lr_PAIR_OFFSET						: LREAL := 70;	// [mm] Delta 1: cups on either side of the flange along the tool's X
	lr_TILT_DIAMETER					: LREAL := 30;	// [mm] Delta 2
	lr_TILT_HEIGHT						: LREAL := 90;	// [mm]
	lr_TILT_ANGLE						: LREAL := 25;	// [deg] about Rx while carrying
	lr_TILT_SPEED						: LREAL := 60;	// [deg/s]
	n_RING_FINGERS						: INT := 5;	// [-] Delta 3
	lr_RING_DIAMETER					: LREAL := 16;	// [mm]
	lr_RING_HEIGHT						: LREAL := 40;	// [mm] reaching down to the belt beside a carried product
	lr_SPREAD_OPEN						: LREAL := 130;	// [mm]
	lr_RING_CLEARANCE					: LREAL := 10;	// [mm] closed fingers: finger radius plus a gap beyond the product's corners
	lr_SPREAD_SPEED						: LREAL := 200;	// [mm/s]
	(* Sequence *)
	n_PHASE_IDLE						: INT := 0;
	n_PHASE_APPROACH					: INT := 1;
	n_PHASE_DESCEND						: INT := 2;
	n_PHASE_LIFT						: INT := 3;
	n_PHASE_TRANSFER					: INT := 4;
	n_PHASE_LOWER						: INT := 5;
	n_PHASE_RELEASE						: INT := 6;
	(* Sequence control *)
	lr_TCP_ACCEL						: LREAL := 20000;	// [mm/s2] Delta 1's TCP acceleration at 100 %
	lr_MISSED_HOLD						: LREAL := 3;	// [s] the missed-product message stays after the last missed product
	udn_RANDOM_A						: UDINT := 1664525;	// [-] the generator's linear congruential pseudo-random numbers
	udn_RANDOM_C						: UDINT := 1013904223;	// [-]
END_VAR

lr_Dt := DEMO_GlobalVar.DEMO_lr_Dt;


(****************************************************************************************************)
(* REGISTRATION (idempotent, every cycle)                                                           *)
(****************************************************************************************************)
fb_Infeed1.m_Register(vio_Manifest := GVL_Visu.stManifest, vi_udn_Id := 1, vi_str_Name := 'Infeed 1');
fb_Infeed2.m_Register(vio_Manifest := GVL_Visu.stManifest, vi_udn_Id := 2, vi_str_Name := 'Infeed 2');
fb_Outfeed.m_Register(vio_Manifest := GVL_Visu.stManifest, vi_udn_Id := 3, vi_str_Name := 'Outfeed');
fb_Delta1.m_Register(vio_Manifest := GVL_Visu.stManifest, vi_udn_Id := 10, vi_str_Name := 'Delta 1');
fb_Delta2.m_Register(vio_Manifest := GVL_Visu.stManifest, vi_udn_Id := 11, vi_str_Name := 'Delta 2');
fb_Delta3.m_Register(vio_Manifest := GVL_Visu.stManifest, vi_udn_Id := 12, vi_str_Name := 'Delta 3');
fb_Vision1.m_Register(vio_Manifest := GVL_Visu.stManifest, vi_udn_Id := 50, vi_str_Name := 'Vision 1');
fb_Barrier2.m_Register(vio_Manifest := GVL_Visu.stManifest, vi_udn_Id := 51, vi_str_Name := 'Light barrier 2');
fb_RejectUnit.m_Register(vio_Manifest := GVL_Visu.stManifest, vi_udn_Id := 60, vi_str_Name := 'Reject unit');
(* What the product mark of a sample means, for the whole PLC. *)
_FC_VisuSetMarkName(vio_Manifest := GVL_Visu.stManifest, vi_un_Mark := un_SAMPLE_MARK, vi_str_Name := 'Sample');


(****************************************************************************************************)
(* CONVEYORS (configuration idempotent, every cycle)                                                *)
(****************************************************************************************************)
(* Infeed 1's program values; its parameter set (Syn_Config) replaces them once the configurator wrote one. *)
Infeed1Default.stPose.fX := 0;
Infeed1Default.stPose.fY := lr_INFEED1_Y;
Infeed1Default.stPose.fZ := DEMO_GlobalConst.DEMO_lr_BELT_Z;
Infeed1Default.nProductTypeCount := UDINT_TO_UINT(udn_TYPE_COUNT);
FOR udn_Type := 1 TO udn_TYPE_COUNT DO
	Infeed1Default.aProductTypes[udn_Type - 1].nId := udn_Type;
	Infeed1Default.aProductTypes[udn_Type - 1].fLength := lr_TYPE_LENGTH[udn_Type];
	Infeed1Default.aProductTypes[udn_Type - 1].fWidth := lr_TYPE_WIDTH[udn_Type];
	Infeed1Default.aProductTypes[udn_Type - 1].fHeight := lr_TYPE_HEIGHT[udn_Type];
	Infeed1Default.aProductTypes[udn_Type - 1].eShape := e_TYPE_SHAPE[udn_Type];
	Infeed1Default.aProductTypes[udn_Type - 1].fCornerRadius := lr_TYPE_CORNER_RADIUS[udn_Type];
END_FOR
fb_Infeed1Param.m_Register(vio_Manifest := GVL_Config.stManifest, vi_udn_Id := fb_Infeed1.m_Id());
fb_Infeed1Param.m_Cycle(vio_Default := Infeed1Default, vio_Set := Infeed1Set, vi_b_ApplyAllowed := TRUE);

FOR n_Belt := 0 TO 2 DO
	CASE n_Belt OF
		0: fb_RefBelt REF= fb_Infeed1;
		1: fb_RefBelt REF= fb_Infeed2; BeltPose := Infeed1Default.stPose; BeltPose.fY := lr_INFEED2_Y;
	ELSE
		fb_RefBelt REF= fb_Outfeed; BeltPose := Infeed1Default.stPose; BeltPose.fY := lr_OUTFEED_Y;
	END_CASE
	fb_RefBelt.m_Configure(vi_lr_Length := lr_BELT_LENGTH, vi_lr_Width := DEMO_GlobalConst.DEMO_lr_BELT_WIDTH);
	(* Infeed 1's pose and product types come with its parameter set (m_PassOn below). *)
	IF n_Belt <> 0 THEN
		fb_RefBelt.m_SetPose(vi_Pose := BeltPose);
		FOR udn_Type := 1 TO udn_TYPE_COUNT DO
			fb_RefBelt.m_SetProductType(vi_udn_Id := udn_Type, vi_lr_Length := lr_TYPE_LENGTH[udn_Type],
				vi_lr_Width := lr_TYPE_WIDTH[udn_Type], vi_lr_Height := lr_TYPE_HEIGHT[udn_Type],
				vi_e_Shape := e_TYPE_SHAPE[udn_Type], vi_lr_CornerRadius := lr_TYPE_CORNER_RADIUS[udn_Type]);
		END_FOR
	END_IF
END_FOR
fb_Infeed1Param.m_PassOn(vio_Visu := fb_Infeed1);
fb_Infeed2.m_SetOriginShift(vi_lr_X := lr_INFEED2_ORIGIN_X, vi_lr_Y := 0, vi_lr_Z := 0);
fb_Outfeed.m_SetOriginShift(vi_lr_X := lr_OUTFEED_ORIGIN_X, vi_lr_Y := 0, vi_lr_Z := 0);

(* Belt travel *)
lr_BeltPosition[0] := lr_BeltPosition[0] + DEMO_GlobalVar.DEMO_lr_Infeed1Speed * lr_Dt;	// ramped by the sequence control
lr_BeltPosition[1] := lr_BeltPosition[1] + lr_INFEED_SPEED * lr_Dt;
lr_BeltPosition[2] := lr_BeltPosition[2] + lr_OUTFEED_SPEED * lr_Dt;
fb_Infeed1.m_SetBeltPosition(lr_BeltPosition[0]);
fb_Infeed2.m_SetBeltPosition(lr_BeltPosition[1]);
fb_Outfeed.m_SetBeltPosition(lr_BeltPosition[2]);


(****************************************************************************************************)
(* DETECTORS (configuration idempotent, every cycle)                                                *)
(****************************************************************************************************)
(* Vision 1's program values; its parameter set (Syn_Config) replaces them once the configurator wrote one. The
   field of view is hardware and stays the program's. *)
Vision1Default.stPose.fX := lr_VISION_X;
Vision1Default.stPose.fY := lr_INFEED1_Y;
Vision1Default.stPose.fZ := DEMO_GlobalConst.DEMO_lr_BELT_Z + lr_VISION_DISTANCE;
Vision1Default.nZoneCount := 1;
Vision1Default.aZones[0].nConveyorId := fb_Infeed1.m_Id();
Vision1Default.aZones[0].fStart := lr_VISION_X - lr_VISION_FIELD / 2;
Vision1Default.aZones[0].fEnd := lr_VISION_X + lr_VISION_FIELD / 2;
Vision1Default.aZones[0].fCcsOffset := lr_VISION_X;
fb_Vision1Param.m_Register(vio_Manifest := GVL_Config.stManifest, vi_udn_Id := fb_Vision1.m_Id());
fb_Vision1Param.m_Cycle(vio_Default := Vision1Default, vio_Set := Vision1Set, vi_b_ApplyAllowed := TRUE);
fb_Vision1.m_Configure(vi_lr_FieldLength := lr_VISION_FIELD, vi_lr_FieldWidth := lr_VISION_FIELD,
	vi_lr_WorkingDistance := lr_VISION_DISTANCE);
fb_Vision1Param.m_PassOn(vio_Visu := fb_Vision1);
(* The head at the right belt edge, its beam across the belt towards +Y. Infeed 2 counts from its end. *)
DetectorPose.fX := lr_BARRIER_X;
DetectorPose.fY := lr_INFEED2_Y - lr_BARRIER_BEAM / 2;
DetectorPose.fZ := DEMO_GlobalConst.DEMO_lr_BELT_Z + lr_BARRIER_HEIGHT;
fb_Barrier2.m_SetPose(vi_Pose := DetectorPose);
fb_Barrier2.m_Configure(vi_lr_BeamLength := lr_BARRIER_BEAM);
fb_Barrier2.m_SetZone(vi_un_Zone := 1, vi_udn_ConveyorId := fb_Infeed2.m_Id(), vi_lr_Start := lr_BARRIER_X - lr_INFEED2_ORIGIN_X,
	vi_lr_End := lr_BARRIER_X - lr_INFEED2_ORIGIN_X, vi_lr_AllocationOffset := 0,
	vi_lr_CcsOffset := lr_BARRIER_X - lr_INFEED2_ORIGIN_X, vi_lr_StartY := 0, vi_lr_EndY := 0);


(****************************************************************************************************)
(* PRODUCT INFEED: Infeed 1 from the product generator, Infeed 2 every lr_SPAWN_INTERVAL             *)
(****************************************************************************************************)
(* Reset accepted by the sequence control: Infeed 1 and Delta 1 start empty, the generator from its seed. *)
IF DEMO_GlobalVar.DEMO_b_Reset THEN
	m_Reset();
END_IF
(* Infeed 1: the generator makes up a detection, the tracking latches it as Vision 1's. *)
IF m_Generate(vo_Detection => Detection) THEN
	m_Track(vi_Detection := Detection);
END_IF
(* Infeed 2: products slightly offset across the belt and turned, latched where the light barrier sees their front
   edge. *)
lr_SinceSpawn2 := lr_SinceSpawn2 + lr_Dt;
IF lr_SinceSpawn2 >= lr_SPAWN_INTERVAL THEN
	lr_SinceSpawn2 := 0;
	udn_Seed := udn_Seed * 1103515245 + 12345;
	lr_Random := UDINT_TO_LREAL(udn_Seed MOD 1000) / 1000.0;
	LatchPose.fY := lr_INFEED2_Y + (lr_Random - 0.5) * 160.0;
	LatchPose.fZ := DEMO_GlobalConst.DEMO_lr_BELT_Z;
	LatchPose.fRz := (UDINT_TO_LREAL((udn_Seed / 1000) MOD 1000) / 1000.0 - 0.5) * 60.0;
	udn_Type := (udn_Seed / 1000000) MOD udn_TYPE_COUNT + 1;
	LatchPose.fX := lr_BARRIER_X - lr_TYPE_LENGTH[udn_Type] / 2;
	IF fb_Infeed2.m_LatchProduct(vi_udn_Id := DEMO_GlobalVar.DEMO_udn_NextId,
		vi_LatchPose := fb_Infeed2.m_McsToBelt(vi_Pose := LatchPose),
		vi_udn_ProductType := udn_Type, vi_lr_LatchBeltPosition := 0, vi_b_UseLatchBeltPosition := FALSE,
		vi_e_State := E_VisuProductState.DETECTED, vi_udn_ClientId := fb_Barrier2.m_Id())
	THEN
		DEMO_GlobalVar.DEMO_udn_NextId := DEMO_GlobalVar.DEMO_udn_NextId + 1;
	END_IF
END_IF


(****************************************************************************************************)
(* ROBOTS: per robot configure it, follow its target, run its sequence and report it                *)
(****************************************************************************************************)
FOR n_Robot := 0 TO 2 DO
	(* Delta 1 runs with the recipe and as fast as its belt, so it halts with it; the others at full speed. *)
	IF n_Robot = 0 THEN
		lr_Step := m_Delta1Step();
	ELSE
		lr_Step := lr_TCP_SPEED * lr_Dt;
	END_IF
	m_Configure();
	m_Target();
	m_Sequence();
	m_Report();
END_FOR


(* The light barrier's beam is interrupted while a product not yet picked covers it. *)
b_BeamInterrupted := FALSE;
un_Index := 0;
WHILE un_Index < fb_Infeed2.m_ProductCount() DO
	fb_Infeed2.m_GetProduct(vi_un_Index := un_Index, vo_Product => Product, vo_Pose => ProductPose);
	ProductPose := fb_Infeed2.m_BeltToMcs(vi_Pose := ProductPose);
	IF Product.eState <> E_VisuProductState.PICKED AND Product.nProductType >= 1 AND Product.nProductType <= udn_TYPE_COUNT
		AND_THEN ABS(ProductPose.fX - lr_BARRIER_X) <= lr_TYPE_LENGTH[Product.nProductType] / 2
	THEN
		b_BeamInterrupted := TRUE;
	END_IF
	un_Index := un_Index + 1;
END_WHILE
fb_Barrier2.m_SetSignal(vi_b_Signal := b_BeamInterrupted);
m_RejectUnit();


(****************************************************************************************************)
(* HOUSEKEEPING                                                                                     *)
(****************************************************************************************************)
m_Missed();
(* Drop register entries some distance beyond the belt end, so "missed" stays visible briefly. *)
fb_Infeed1.m_RemoveProductsBeyond(lr_BELT_LENGTH + DEMO_GlobalConst.DEMO_lr_REMOVE_BEYOND_END);
fb_Infeed2.m_RemoveProductsBeyond(lr_BELT_LENGTH + DEMO_GlobalConst.DEMO_lr_REMOVE_BEYOND_END);
fb_Outfeed.m_RemoveProductsBeyond(lr_BELT_LENGTH + DEMO_GlobalConst.DEMO_lr_REMOVE_BEYOND_END);

(****************************************************************************************************<br>
© Syntegon Group.<br>
All rights reserved, also regarding any disposal, exploitation, reproduction, editing, distribution,<br>
as well as in the event of applications for industrial property rights.<br>
*****************************************************************************************************<br>
DESCRIPTION:<br>
Looks for a detected product in the allocation area of Delta n_Robot and assigns it. Delta 1 serves infeed 1,<br>
Delta 2 infeed 2, Delta 3 takes what both leave. TRUE if a product was assigned.<br>
****************************************************************************************************)
METHOD PRIVATE m_Allocate : BOOL
VAR
	TempStart							: ST_VisuPlanarPose;	// start of Delta 1's allocation area, belt coordinates, then MCS
	TempEnd								: ST_VisuPlanarPose;	// its end, belt coordinates, then MCS
END_VAR
FOR n_Belt := 0 TO 1 DO
	IF n_Belt = 0 THEN
		fb_RefBelt REF= fb_Infeed1;
	ELSE
		fb_RefBelt REF= fb_Infeed2;
	END_IF
	(* Where the robot allocates on this infeed: around its base, Delta 1 on infeed 1 in the pick zone of its parameter
	   set (belt coordinates to MCS X: infeed 1 runs along +X). *)
	lr_AllocStart := lr_BaseX - lr_PICK_HALF_ZONE;
	lr_AllocEnd := lr_BaseX + lr_PICK_HALF_ZONE - lr_ALLOCATION_OFFSET;
	IF n_Robot = 0 AND n_Belt = 0 AND fb_Delta1Param.m_ZoneCount() >= 1 THEN
		Zone := fb_Delta1Param.m_Zone(vi_un_Zone := 1);
		TempStart.fX := MIN(Zone.fStart, Zone.fEnd);
		TempEnd.fX := MAX(Zone.fStart, Zone.fEnd) - Zone.fAllocationOffset;
		TempStart := fb_Infeed1.m_BeltToMcs(vi_Pose := TempStart);
		TempEnd := fb_Infeed1.m_BeltToMcs(vi_Pose := TempEnd);
		lr_AllocStart := TempStart.fX;
		lr_AllocEnd := TempEnd.fX;
	END_IF
	un_Index := 0;
	(* Nobody takes a product from Infeed 1 while it stands: the machine is stopping or stopped. *)
	IF (n_Robot = 0 AND n_Belt = 1) OR (n_Robot = 1 AND n_Belt = 0)
	OR (n_Belt = 0 AND DEMO_GlobalVar.DEMO_lr_Infeed1Speed = 0)
	THEN
		un_Index := fb_RefBelt.m_ProductCount();
	END_IF
	WHILE udn_TargetId[n_Robot] = 0 AND un_Index < fb_RefBelt.m_ProductCount() DO
		fb_RefBelt.m_GetProduct(vi_un_Index := un_Index, vo_Product => Product, vo_Pose => ProductPose);
		ProductPose := fb_RefBelt.m_BeltToMcs(vi_Pose := ProductPose);
		(* Delta 1 adds only a product of the type it already carries: both cups hang at the same height. *)
		IF Product.eState = E_VisuProductState.DETECTED
		AND (n_Robot <> 0 OR n_HeldCount[n_Robot] = 0 OR Product.nProductType = udn_HeldType[n_Robot, 0])
		AND ProductPose.fX >= lr_AllocStart
		AND ProductPose.fX <= lr_AllocEnd
		THEN
			fb_RefBelt.m_SetProductState(vi_udn_Id := Product.nId, vi_e_State := E_VisuProductState.ASSIGNED,
				vi_udn_ClientId := fb_RefRobot.m_Id(), vi_udn_MoverId := 0, vi_udn_FingerId := 0);
			udn_TargetId[n_Robot] := Product.nId;
			n_TargetBelt[n_Robot] := n_Belt;
			n_Phase[n_Robot] := n_PHASE_APPROACH;
		END_IF
		un_Index := un_Index + 1;
	END_WHILE
END_FOR
m_Allocate := udn_TargetId[n_Robot] <> 0;
END_METHOD

(****************************************************************************************************<br>
© Syntegon Group.<br>
All rights reserved, also regarding any disposal, exploitation, reproduction, editing, distribution,<br>
as well as in the event of applications for industrial property rights.<br>
*****************************************************************************************************<br>
DESCRIPTION:<br>
Selects Delta n_Robot into fb_RefRobot and configures it (idempotent): base, gripper with the fingers' places<br>
on the flange, working area, limit area, TCP limit area and zones. Initialises its TCP once.<br>
****************************************************************************************************)
METHOD PRIVATE m_Configure : BOOL
VAR
	lr_TempAngle						: LREAL;	// [deg] a ring finger's place around the flange
END_VAR
CASE n_Robot OF
	0: fb_RefRobot REF= fb_Delta1;
	1: fb_RefRobot REF= fb_Delta2;
ELSE
	fb_RefRobot REF= fb_Delta3;
END_CASE
lr_BaseX := lr_ROBOT1_X + INT_TO_LREAL(n_Robot) * lr_ROBOT_PITCH;


(****************************************************************************************************
PROGRAM VALUES: base, areas and zones
****************************************************************************************************)
RobotDefault.stPose.fX := lr_BaseX;
RobotDefault.stPose.fY := lr_ROBOT_Y;
RobotDefault.stPose.fZ := lr_ROBOT_Z;
(* The robot's coordinate system sits in its working plane, 900 mm below the base. *)
RobotDefault.stOriginShift.fX := 0;
RobotDefault.stOriginShift.fY := 0;
RobotDefault.stOriginShift.fZ := -900;
RobotDefault.stWorkingArea.fRadius := 750;
RobotDefault.stWorkingArea.fZMin := -1300;
RobotDefault.stWorkingArea.fZMax := -700;
RobotDefault.stWorkingArea.fConeHeight := 200;
RobotDefault.stWorkingArea.fConeBottomRadius := 450;
(* Neighbouring robots share the space between them: each one is limited to half the robot pitch. *)
RobotDefault.stLimitArea.fXMin := -lr_ROBOT_PITCH / 2;
RobotDefault.stLimitArea.fXMax := lr_ROBOT_PITCH / 2;
RobotDefault.stLimitArea.fYMin := -750;
RobotDefault.stLimitArea.fYMax := 750;
RobotDefault.stLimitArea.fZMin := -1500;
RobotDefault.stLimitArea.fZMax := -700;
RobotDefault.stLimitArea.bActive := TRUE;
(* Around the TCP: gripper and product below the flange. It lights up when it reaches into a neighbour's limit
   area or out of the robot's own. *)
RobotDefault.stTcpLimitArea.fXMin := -80;
RobotDefault.stTcpLimitArea.fXMax := 80;
RobotDefault.stTcpLimitArea.fYMin := -80;
RobotDefault.stTcpLimitArea.fYMax := 80;
RobotDefault.stTcpLimitArea.fZMin := -100;
RobotDefault.stTcpLimitArea.fZMax := 20;
RobotDefault.stTcpLimitArea.bActive := TRUE;
(* The robot's conveyor coordinate system lies under its base on every belt. *)
RobotDefault.nZoneCount := 3;
RobotDefault.aZones[0].nConveyorId := fb_Infeed1.m_Id();
RobotDefault.aZones[0].fStart := lr_BaseX - lr_PICK_HALF_ZONE;
RobotDefault.aZones[0].fEnd := lr_BaseX + lr_PICK_HALF_ZONE;
RobotDefault.aZones[0].fAllocationOffset := lr_ALLOCATION_OFFSET;
RobotDefault.aZones[0].fCcsOffset := lr_BaseX;
RobotDefault.aZones[0].fStartY := -lr_PICK_HALF_LANE;
RobotDefault.aZones[0].fEndY := lr_PICK_HALF_LANE;
RobotDefault.aZones[1].nConveyorId := fb_Infeed2.m_Id();
RobotDefault.aZones[1].fStart := lr_BaseX - lr_PICK_HALF_ZONE - lr_INFEED2_ORIGIN_X;
RobotDefault.aZones[1].fEnd := lr_BaseX + lr_PICK_HALF_ZONE - lr_INFEED2_ORIGIN_X;
RobotDefault.aZones[1].fAllocationOffset := lr_ALLOCATION_OFFSET;
RobotDefault.aZones[1].fCcsOffset := lr_BaseX - lr_INFEED2_ORIGIN_X;
RobotDefault.aZones[1].fStartY := -lr_PICK_HALF_LANE;
RobotDefault.aZones[1].fEndY := lr_PICK_HALF_LANE;
RobotDefault.aZones[2].nConveyorId := fb_Outfeed.m_Id();
RobotDefault.aZones[2].fStart := lr_BaseX - lr_PLACE_HALF_ZONE - lr_OUTFEED_ORIGIN_X;
RobotDefault.aZones[2].fEnd := lr_BaseX + lr_PLACE_HALF_ZONE - lr_OUTFEED_ORIGIN_X;
RobotDefault.aZones[2].fAllocationOffset := 0;
RobotDefault.aZones[2].fCcsOffset := lr_BaseX - lr_OUTFEED_ORIGIN_X;
RobotDefault.aZones[2].fStartY := 0;
RobotDefault.aZones[2].fEndY := 0;


(****************************************************************************************************
GRIPPER: the fingers and their places on the flange at rest (ADR 0018); the demo reports their live poses
****************************************************************************************************)
CASE n_Robot OF
	0:
		(* Two suction cups on either side of the flange along its X. *)
		n_FingerCount := 2;
		FOR n_Finger := 1 TO 2 DO
			RobotDefault.aFingers[n_Finger - 1].fDiameter := DEMO_GlobalConst.DEMO_lr_CUP_DIAMETER;
			RobotDefault.aFingers[n_Finger - 1].fHeight := DEMO_GlobalConst.DEMO_lr_CUP_HEIGHT;
			RobotDefault.aFingers[n_Finger - 1].stOffset.fX := SEL(n_Finger = 1, -lr_PAIR_OFFSET, lr_PAIR_OFFSET);
			RobotDefault.aFingers[n_Finger - 1].stOffset.fY := 0;
			RobotDefault.aFingers[n_Finger - 1].stOffset.fRz := 0;
		END_FOR
	1:
		(* One finger at the flange centre. *)
		n_FingerCount := 1;
		RobotDefault.aFingers[0].fDiameter := lr_TILT_DIAMETER;
		RobotDefault.aFingers[0].fHeight := lr_TILT_HEIGHT;
		RobotDefault.aFingers[0].stOffset.fX := 0;
		RobotDefault.aFingers[0].stOffset.fY := 0;
		RobotDefault.aFingers[0].stOffset.fRz := 0;
ELSE
	(* A ring of fingers around the flange, open, each turned to face the centre. *)
	n_FingerCount := n_RING_FINGERS;
	FOR n_Finger := 1 TO n_RING_FINGERS DO
		lr_TempAngle := 360.0 * INT_TO_LREAL(n_Finger - 1) / INT_TO_LREAL(n_RING_FINGERS);
		RobotDefault.aFingers[n_Finger - 1].fDiameter := lr_RING_DIAMETER;
		RobotDefault.aFingers[n_Finger - 1].fHeight := lr_RING_HEIGHT;
		RobotDefault.aFingers[n_Finger - 1].stOffset.fX := lr_SPREAD_OPEN * COS(lr_TempAngle * VISU_GlobalConst.VISU_lr_DEG_TO_RAD);
		RobotDefault.aFingers[n_Finger - 1].stOffset.fY := lr_SPREAD_OPEN * SIN(lr_TempAngle * VISU_GlobalConst.VISU_lr_DEG_TO_RAD);
		RobotDefault.aFingers[n_Finger - 1].stOffset.fRz := lr_TempAngle;
	END_FOR
END_CASE
RobotDefault.nFingerCount := INT_TO_UINT(n_FingerCount);

(* Delta 1 runs with its parameter set (Syn_Config) once the configurator wrote one, also its pick logic. The
   program values are complete only here: RobotDefault serves all three robots. *)
IF n_Robot = 0 THEN
	fb_Delta1Param.m_Register(vio_Manifest := GVL_Config.stManifest, vi_udn_Id := fb_Delta1.m_Id());
	fb_Delta1Param.m_Cycle(vio_Default := RobotDefault, vio_Set := Delta1Set, vi_b_ApplyAllowed := TRUE);
	BasePose := fb_Delta1Param.m_Pose();
	lr_BaseX := BasePose.fX;
ELSE
	BasePose := RobotDefault.stPose;
END_IF
fb_RefRobot.m_Configure(vi_lr_BaseRadius := 200, vi_lr_EffectorRadius := 50,
	vi_lr_UpperArmLength := 400, vi_lr_LowerArmLength := 1000);

(* Delta 1 gets its fingers with its parameter set (m_PassOn below), the others here. *)
IF n_Robot <> 0 THEN
	FOR n_Finger := 1 TO n_FingerCount DO
		fb_RefRobot.m_SetFinger(vi_un_Finger := INT_TO_UINT(n_Finger), vi_lr_Diameter := RobotDefault.aFingers[n_Finger - 1].fDiameter,
			vi_lr_Height := RobotDefault.aFingers[n_Finger - 1].fHeight);
		fb_RefRobot.m_SetFingerOffset(vi_un_Finger := INT_TO_UINT(n_Finger),
			vi_lr_X := RobotDefault.aFingers[n_Finger - 1].stOffset.fX, vi_lr_Y := RobotDefault.aFingers[n_Finger - 1].stOffset.fY,
			vi_lr_Z := RobotDefault.aFingers[n_Finger - 1].stOffset.fZ, vi_lr_Rz := RobotDefault.aFingers[n_Finger - 1].stOffset.fRz);
	END_FOR
END_IF


(****************************************************************************************************
AREAS AND ZONES: Delta 1's from its parameter set, the others' program values
****************************************************************************************************)
IF n_Robot = 0 THEN
	fb_Delta1Param.m_PassOn(vio_Visu := fb_RefRobot);
ELSE
	fb_RefRobot.m_SetPose(vi_Pose := BasePose);
	fb_RefRobot.m_SetWorkingArea(vi_lr_Radius := RobotDefault.stWorkingArea.fRadius,
		vi_lr_ZMin := RobotDefault.stWorkingArea.fZMin, vi_lr_ZMax := RobotDefault.stWorkingArea.fZMax,
		vi_lr_ConeHeight := RobotDefault.stWorkingArea.fConeHeight,
		vi_lr_ConeBottomRadius := RobotDefault.stWorkingArea.fConeBottomRadius);
	fb_RefRobot.m_SetLimitArea(vi_lr_XMin := RobotDefault.stLimitArea.fXMin, vi_lr_XMax := RobotDefault.stLimitArea.fXMax,
		vi_lr_YMin := RobotDefault.stLimitArea.fYMin, vi_lr_YMax := RobotDefault.stLimitArea.fYMax,
		vi_lr_ZMin := RobotDefault.stLimitArea.fZMin, vi_lr_ZMax := RobotDefault.stLimitArea.fZMax);
	fb_RefRobot.m_SetTcpLimitArea(vi_lr_XMin := RobotDefault.stTcpLimitArea.fXMin,
		vi_lr_XMax := RobotDefault.stTcpLimitArea.fXMax, vi_lr_YMin := RobotDefault.stTcpLimitArea.fYMin,
		vi_lr_YMax := RobotDefault.stTcpLimitArea.fYMax, vi_lr_ZMin := RobotDefault.stTcpLimitArea.fZMin,
		vi_lr_ZMax := RobotDefault.stTcpLimitArea.fZMax);
	FOR n_Zone := 1 TO UINT_TO_INT(RobotDefault.nZoneCount) DO
		fb_RefRobot.m_SetZone(vi_un_Zone := INT_TO_UINT(n_Zone), vi_udn_ConveyorId := RobotDefault.aZones[n_Zone - 1].nConveyorId,
			vi_lr_Start := RobotDefault.aZones[n_Zone - 1].fStart, vi_lr_End := RobotDefault.aZones[n_Zone - 1].fEnd,
			vi_lr_AllocationOffset := RobotDefault.aZones[n_Zone - 1].fAllocationOffset,
			vi_lr_CcsOffset := RobotDefault.aZones[n_Zone - 1].fCcsOffset,
			vi_lr_StartY := RobotDefault.aZones[n_Zone - 1].fStartY, vi_lr_EndY := RobotDefault.aZones[n_Zone - 1].fEndY);
	END_FOR
	fb_RefRobot.m_SetOriginShift(vi_lr_X := RobotDefault.stOriginShift.fX, vi_lr_Y := RobotDefault.stOriginShift.fY,
		vi_lr_Z := RobotDefault.stOriginShift.fZ);
END_IF

(* Start position of the TCP *)
IF NOT b_TcpInitialised[n_Robot] THEN
	Tcp[n_Robot].fX := lr_BaseX;
	Tcp[n_Robot].fY := lr_ROBOT_Y;
	Tcp[n_Robot].fZ := lr_ROBOT_Z - 900;
	b_TcpInitialised[n_Robot] := TRUE;
END_IF
m_Configure := TRUE;
END_METHOD

(****************************************************************************************************<br>
© Syntegon Group.<br>
All rights reserved, also regarding any disposal, exploitation, reproduction, editing, distribution,<br>
as well as in the event of applications for industrial property rights.<br>
*****************************************************************************************************<br>
DESCRIPTION:<br>
Delta 1's TCP travel this cycle: its speed ramps with the recipe's acceleration (% of lr_TCP_ACCEL) towards the<br>
recipe's speed (% of lr_TCP_SPEED), scaled by how far Infeed 1 is at its recipe speed, so the robot slows down and<br>
halts with its belt when the machine stops.<br>
****************************************************************************************************)
METHOD PRIVATE m_Delta1Step : LREAL
VAR
	lr_TempBeltShare					: LREAL;	// [-] Infeed 1's speed of its recipe speed, 0..1
	lr_TempTarget						: LREAL;	// [mm/s]
	lr_TempChange						: LREAL;	// [mm/s] at most this cycle
END_VAR
lr_TempBeltShare := LIMIT(0.0, DEMO_GlobalVar.DEMO_lr_Infeed1Speed / MAX(DEMO_GlobalVar.DEMO_Recipe.lr_BeltSpeed, 1.0), 1.0);
lr_TempTarget := lr_TCP_SPEED * DEMO_GlobalVar.DEMO_Recipe.lr_RobotSpeed / 100.0 * lr_TempBeltShare;
lr_TempChange := lr_TCP_ACCEL * DEMO_GlobalVar.DEMO_Recipe.lr_RobotAccel / 100.0 * lr_Dt;
lr_Delta1Speed := _FC_DemoApproach(lr_Delta1Speed, lr_TempTarget, lr_TempChange);
m_Delta1Step := lr_Delta1Speed * lr_Dt;
END_METHOD

(****************************************************************************************************<br>
© Syntegon Group.<br>
All rights reserved, also regarding any disposal, exploitation, reproduction, editing, distribution,<br>
as well as in the event of applications for industrial property rights.<br>
*****************************************************************************************************<br>
DESCRIPTION:<br>
Pose of a Delta's finger frame (centre of its top face), absolute in the MCS, from the robot's TCP (the flange)<br>
and its tool state:<br>
- Delta 1: two cups on either side of the flange at lr_PAIR_OFFSET along the tool's X, turned by lr_ToolRz.<br>
- Delta 2: one finger at the flange, turned by lr_ToolRz and tilted about its own X by lr_TiltRx.<br>
- Delta 3: n_RING_FINGERS fingers on a circle of radius lr_Spread around the flange, each facing outwards.<br>
****************************************************************************************************)
METHOD PRIVATE m_FingerPose : ST_VisuPose
VAR_INPUT
	vi_n_Robot							: INT;	// [-] 0..2
	vi_n_Finger							: INT;	// [-] 1-based
END_VAR
VAR
	lr_TempRz							: LREAL;	// [deg]
	lr_TempRadius						: LREAL;	// [mm] finger distance from the flange
END_VAR
m_FingerPose.fX := Tcp[vi_n_Robot].fX;
m_FingerPose.fY := Tcp[vi_n_Robot].fY;
m_FingerPose.fZ := Tcp[vi_n_Robot].fZ;
m_FingerPose.fRx := 0;
m_FingerPose.fRy := 0;
lr_TempRz := lr_ToolRz[vi_n_Robot];
lr_TempRadius := 0;
CASE vi_n_Robot OF
	0:
		(* Finger 1 along the tool's +X, finger 2 along its -X. *)
		lr_TempRadius := SEL(vi_n_Finger = 1, -lr_PAIR_OFFSET, lr_PAIR_OFFSET);
	1:
		m_FingerPose.fRx := lr_TiltRx;
	2:
		lr_TempRz := lr_ToolRz[vi_n_Robot] + 360.0 / INT_TO_LREAL(n_RING_FINGERS) * INT_TO_LREAL(vi_n_Finger - 1);
		lr_TempRadius := lr_Spread;
END_CASE
m_FingerPose.fX := m_FingerPose.fX + lr_TempRadius * COS(lr_TempRz * VISU_GlobalConst.VISU_lr_DEG_TO_RAD);
m_FingerPose.fY := m_FingerPose.fY + lr_TempRadius * SIN(lr_TempRz * VISU_GlobalConst.VISU_lr_DEG_TO_RAD);
m_FingerPose.fRz := lr_TempRz;
END_METHOD

(****************************************************************************************************<br>
© Syntegon Group.<br>
All rights reserved, also regarding any disposal, exploitation, reproduction, editing, distribution,<br>
as well as in the event of applications for industrial property rights.<br>
*****************************************************************************************************<br>
DESCRIPTION:<br>
The product generator on Infeed 1 before Vision 1, from the recipe's product pattern: a place every so many mm of<br>
belt travel (the rate at the recipe's belt speed, so the pattern keeps its spacing while the belt ramps or stands),<br>
a share of the places left empty, each product of a type of the type mix and, by the pattern, in one of the lanes<br>
at random (Lanes) or in the one lane, scattered along and across the belt (never off it) and turned (Scattered).<br>
It makes up a raw detection as a vision system would report<br>
it: the product's pose, the belt position at that moment, its type; m_Track latches it. A new seed, or a reset,<br>
starts the numbers again: the same seed gives the same products.<br>
*****************************************************************************************************<br>
OUTPUT VALUES:<br>
TRUE in the cycle it made up a detection (vo_Detection).<br>
****************************************************************************************************)
METHOD PRIVATE m_Generate : BOOL
VAR_OUTPUT
	vo_Detection						: TVisuDemo_Detection;
END_VAR
VAR
	lr_TempSpacing						: LREAL;	// [mm] belt travel between the generator's places
	dn_TempLanes						: DINT;	// [-]
	lr_TempY							: LREAL;	// [mm] across the belt from its middle
	lr_TempHalfWidth					: LREAL;	// [mm] how far from the middle a product may lie
	lr_TempScatter						: LREAL;	// [-] 1: the pattern scatters (Scattered), 0: not (Lanes)
	TempLens							: ST_VisuPose;	// Vision 1's effective pose, MCS
	TempMcs								: ST_VisuPlanarPose;	// the lens as a planar pose, MCS
	TempBelt							: ST_VisuPlanarPose;	// the detection in Infeed 1's coordinate system
END_VAR
m_Generate := FALSE;
IF DEMO_GlobalVar.DEMO_Recipe.dn_Seed <> dn_GenSeed THEN
	dn_GenSeed := DEMO_GlobalVar.DEMO_Recipe.dn_Seed;
	udn_GenRandom := DINT_TO_UDINT(dn_GenSeed);
	lr_GenTravel := 0;
	un_Vision1Latches := 0;
END_IF
IF NOT DEMO_GlobalVar.DEMO_Recipe.b_Feed OR DEMO_GlobalVar.DEMO_Recipe.lr_Rate <= 0 THEN
	RETURN;
END_IF

(* A place every lr_TempSpacing of belt travel; a shorter spacing (a higher rate) starts from the next place, so the
   travel gathered before never pours out at once. *)
lr_TempSpacing := MAX(DEMO_GlobalVar.DEMO_Recipe.lr_BeltSpeed, 1) * 60.0 / DEMO_GlobalVar.DEMO_Recipe.lr_Rate;
lr_GenTravel := MIN(lr_GenTravel + DEMO_GlobalVar.DEMO_lr_Infeed1Speed * lr_Dt, lr_TempSpacing);
IF lr_GenTravel < lr_TempSpacing THEN
	RETURN;
END_IF
lr_GenTravel := 0;
IF m_Random() * 100.0 < DEMO_GlobalVar.DEMO_Recipe.lr_GapShare THEN
	RETURN;	// a gap
END_IF

(* Its lane, type and scatter, on the belt: the pattern Lanes puts it into one of its lanes unscattered, Scattered
   into the one lane, scattered. Both draw the same numbers, so a seed gives the same products in either. *)
IF DEMO_GlobalVar.DEMO_Recipe.b_PatternLanes THEN
	dn_TempLanes := LIMIT(1, DEMO_GlobalVar.DEMO_Recipe.dn_Lanes, 4);
	lr_TempScatter := 0;
ELSE
	dn_TempLanes := 1;
	lr_TempScatter := 1;
END_IF
lr_TempY := (DINT_TO_LREAL(m_RandomIndex(vi_dn_Count := dn_TempLanes)) - DINT_TO_LREAL(dn_TempLanes - 1) / 2.0)
	* DEMO_GlobalVar.DEMO_Recipe.lr_LanePitch
	+ (m_Random() * 2.0 - 1.0) * DEMO_GlobalVar.DEMO_Recipe.lr_ScatterY * lr_TempScatter;
lr_TempHalfWidth := DEMO_GlobalConst.DEMO_lr_BELT_WIDTH / 2.0 - 50.0;
CASE DEMO_GlobalVar.DEMO_Recipe.dn_TypeMix OF
	1: vo_Detection.udn_ProductType := 1 + DINT_TO_UDINT(m_RandomIndex(vi_dn_Count := 2));	// boxes: 1, 2
	2: vo_Detection.udn_ProductType := 3 + DINT_TO_UDINT(m_RandomIndex(vi_dn_Count := 2));	// round: the can, the oval
ELSE
	vo_Detection.udn_ProductType := 1 + DINT_TO_UDINT(m_RandomIndex(vi_dn_Count := UDINT_TO_DINT(udn_TYPE_COUNT)));
END_CASE
(* On Infeed 1 under Vision 1's lens, in the belt's coordinates; the camera reports it in the MCS. *)
TempLens := fb_Vision1Param.m_Pose();
TempMcs.fX := TempLens.fX;
TempMcs.fY := TempLens.fY;
TempMcs.fZ := TempLens.fZ;
TempBelt := fb_Infeed1.m_McsToBelt(vi_Pose := TempMcs);
TempBelt.fX := TempBelt.fX + (m_Random() * 2.0 - 1.0) * DEMO_GlobalVar.DEMO_Recipe.lr_ScatterX * lr_TempScatter;
TempBelt.fY := LIMIT(-lr_TempHalfWidth, lr_TempY, lr_TempHalfWidth);
TempBelt.fZ := 0;
TempBelt.fRz := (m_Random() * 2.0 - 1.0) * DEMO_GlobalVar.DEMO_Recipe.lr_ScatterRz * lr_TempScatter;
vo_Detection.Pose := fb_Infeed1.m_BeltToMcs(vi_Pose := TempBelt);
vo_Detection.lr_BeltPosition := lr_BeltPosition[0];
m_Generate := TRUE;
END_METHOD

(****************************************************************************************************<br>
© Syntegon Group.<br>
All rights reserved, also regarding any disposal, exploitation, reproduction, editing, distribution,<br>
as well as in the event of applications for industrial property rights.<br>
*****************************************************************************************************<br>
DESCRIPTION:<br>
MCS offset from a Delta's TCP (the flange) to the grip point of one of its fingers, the centre of the finger's<br>
bottom face: where a carried product's top touches. vi_n_Finger = 0 is the flange itself.<br>
****************************************************************************************************)
METHOD PRIVATE m_GripOffset : ST_VisuPosition
VAR_INPUT
	vi_n_Robot							: INT;	// [-] 0..2
	vi_n_Finger							: INT;	// [-] 1-based, 0 = flange
END_VAR
VAR
	TempTop								: ST_VisuPose;
	lr_TempHeight						: LREAL;	// [mm]
	lr_TempRx							: LREAL;	// [rad]
	lr_TempRz							: LREAL;	// [rad]
END_VAR
IF vi_n_Finger = 0 THEN
	RETURN;
END_IF
CASE vi_n_Robot OF
	0: lr_TempHeight := DEMO_GlobalConst.DEMO_lr_CUP_HEIGHT;
	1: lr_TempHeight := lr_TILT_HEIGHT;
ELSE
	lr_TempHeight := lr_RING_HEIGHT;
END_CASE
TempTop := m_FingerPose(vi_n_Robot := vi_n_Robot, vi_n_Finger := vi_n_Finger);
lr_TempRx := TempTop.fRx * VISU_GlobalConst.VISU_lr_DEG_TO_RAD;
lr_TempRz := TempTop.fRz * VISU_GlobalConst.VISU_lr_DEG_TO_RAD;
(* Rz(rz) * Rx(rx) * (0, 0, -height): the finger's local -Z in the MCS. *)
m_GripOffset.fX := TempTop.fX - Tcp[vi_n_Robot].fX - lr_TempHeight * SIN(lr_TempRx) * SIN(lr_TempRz);
m_GripOffset.fY := TempTop.fY - Tcp[vi_n_Robot].fY + lr_TempHeight * SIN(lr_TempRx) * COS(lr_TempRz);
m_GripOffset.fZ := TempTop.fZ - Tcp[vi_n_Robot].fZ - lr_TempHeight * COS(lr_TempRx);
END_METHOD

(****************************************************************************************************<br>
© Syntegon Group.<br>
All rights reserved, also regarding any disposal, exploitation, reproduction, editing, distribution,<br>
as well as in the event of applications for industrial property rights.<br>
*****************************************************************************************************<br>
DESCRIPTION:<br>
Whether a product passed Infeed 1's end unpicked (still DETECTED or ASSIGNED): it raises the machine message<br>
'Product missed' (P_VisuDemoMachine), which stays lr_MISSED_HOLD after the last one.<br>
*****************************************************************************************************<br>
OUTPUT VALUES:<br>
TRUE while a missed product is beyond the belt end.<br>
****************************************************************************************************)
METHOD PRIVATE m_Missed : BOOL
VAR
	un_TempIndex						: UINT;
	TempProduct							: ST_VisuProduct;
	TempPose							: ST_VisuPlanarPose;
END_VAR
m_Missed := FALSE;
un_TempIndex := 0;
WHILE un_TempIndex < fb_Infeed1.m_ProductCount() DO
	fb_Infeed1.m_GetProduct(vi_un_Index := un_TempIndex, vo_Product => TempProduct, vo_Pose => TempPose);
	(* Beyond the belt end, along the belt as m_RemoveProductsBeyond counts. *)
	IF (TempProduct.eState = E_VisuProductState.DETECTED OR TempProduct.eState = E_VisuProductState.ASSIGNED)
	AND TempPose.fX > lr_BELT_LENGTH
	THEN
		m_Missed := TRUE;
	END_IF
	un_TempIndex := un_TempIndex + 1;
END_WHILE
IF m_Missed THEN
	lr_MissedLeft := lr_MISSED_HOLD;
ELSE
	lr_MissedLeft := MAX(0.0, lr_MissedLeft - lr_Dt);
END_IF
DEMO_GlobalVar.DEMO_b_Infeed1Missed := lr_MissedLeft > 0;
END_METHOD

(****************************************************************************************************<br>
© Syntegon Group.<br>
All rights reserved, also regarding any disposal, exploitation, reproduction, editing, distribution,<br>
as well as in the event of applications for industrial property rights.<br>
*****************************************************************************************************<br>
DESCRIPTION:<br>
Moves a TCP towards a target by at most vi_lr_MaxStep. TRUE once the target is reached.<br>
****************************************************************************************************)
METHOD PRIVATE m_MoveToward : BOOL
VAR_IN_OUT
	vio_Tcp								: ST_VisuPosition;
END_VAR
VAR_INPUT
	vi_lr_TargetX						: LREAL;	// [mm]
	vi_lr_TargetY						: LREAL;	// [mm]
	vi_lr_TargetZ						: LREAL;	// [mm]
	vi_lr_MaxStep						: LREAL;	// [mm]
END_VAR
VAR
	lr_TempDx							: LREAL;	// [mm]
	lr_TempDy							: LREAL;	// [mm]
	lr_TempDz							: LREAL;	// [mm]
	lr_TempDist							: LREAL;	// [mm]
END_VAR
lr_TempDx := vi_lr_TargetX - vio_Tcp.fX;
lr_TempDy := vi_lr_TargetY - vio_Tcp.fY;
lr_TempDz := vi_lr_TargetZ - vio_Tcp.fZ;
lr_TempDist := SQRT(lr_TempDx * lr_TempDx + lr_TempDy * lr_TempDy + lr_TempDz * lr_TempDz);
IF lr_TempDist <= vi_lr_MaxStep THEN
	vio_Tcp.fX := vi_lr_TargetX;
	vio_Tcp.fY := vi_lr_TargetY;
	vio_Tcp.fZ := vi_lr_TargetZ;
	m_MoveToward := TRUE;
ELSE
	vio_Tcp.fX := vio_Tcp.fX + lr_TempDx / lr_TempDist * vi_lr_MaxStep;
	vio_Tcp.fY := vio_Tcp.fY + lr_TempDy / lr_TempDist * vi_lr_MaxStep;
	vio_Tcp.fZ := vio_Tcp.fZ + lr_TempDz / lr_TempDist * vi_lr_MaxStep;
	m_MoveToward := FALSE;
END_IF
END_METHOD

(****************************************************************************************************<br>
© Syntegon Group.<br>
All rights reserved, also regarding any disposal, exploitation, reproduction, editing, distribution,<br>
as well as in the event of applications for industrial property rights.<br>
*****************************************************************************************************<br>
DESCRIPTION:<br>
The product generator's next pseudo-random number in 0..1 (below 1): a linear congruential generator, so the same<br>
seed always gives the same numbers.<br>
****************************************************************************************************)
METHOD PRIVATE m_Random : LREAL
udn_GenRandom := udn_GenRandom * udn_RANDOM_A + udn_RANDOM_C;
(* The upper 24 bits: the lower ones of such a generator repeat soon. *)
m_Random := UDINT_TO_LREAL(SHR(udn_GenRandom, 8)) / 16777216.0;
END_METHOD

(****************************************************************************************************<br>
© Syntegon Group.<br>
All rights reserved, also regarding any disposal, exploitation, reproduction, editing, distribution,<br>
as well as in the event of applications for industrial property rights.<br>
*****************************************************************************************************<br>
DESCRIPTION:<br>
One of vi_dn_Count values 0..vi_dn_Count-1, each as likely, from the generator's next pseudo-random number.<br>
****************************************************************************************************)
METHOD PRIVATE m_RandomIndex : DINT
VAR_INPUT
	vi_dn_Count							: DINT;	// [-] at least 1
END_VAR
m_RandomIndex := LIMIT(0, TRUNC(m_Random() * DINT_TO_LREAL(vi_dn_Count)), MAX(vi_dn_Count, 1) - 1);
END_METHOD

(****************************************************************************************************<br>
© Syntegon Group.<br>
All rights reserved, also regarding any disposal, exploitation, reproduction, editing, distribution,<br>
as well as in the event of applications for industrial property rights.<br>
*****************************************************************************************************<br>
DESCRIPTION:<br>
Reject unit at the right edge of the outfeed: describes its housing and pusher and its zone, a line across<br>
the belt at lr_REJECT_X. Every un_REJECT_EVERY-th product passing it is set REJECTED by the reject unit;<br>
the pusher lights up and the product leaves the register after lr_REJECT_PUSH_TIME.<br>
****************************************************************************************************)
METHOD PRIVATE m_RejectUnit : BOOL
VAR
	TempPose							: ST_VisuPose;
	TempProduct							: ST_VisuProduct;
	TempProductPose						: ST_VisuPlanarPose;
	un_TempIndex						: UINT;
END_VAR
VAR CONSTANT
	lr_GAP								: LREAL := 30;	// [mm] between the belt edge and the pusher's back
	lr_HOUSING_LENGTH					: LREAL := 160;	// [mm] along the belt
	lr_HOUSING_WIDTH					: LREAL := 140;	// [mm]
	lr_HOUSING_ABOVE_BELT				: LREAL := 120;	// [mm] its top above the belt surface
	lr_PUSHER_LENGTH					: LREAL := 120;	// [mm] along the belt
	lr_PUSHER_WIDTH						: LREAL := 30;	// [mm]
	lr_PUSHER_HEIGHT					: LREAL := 50;	// [mm]
	lr_PUSHER_ABOVE_BELT				: LREAL := 10;	// [mm] its bottom above the belt surface
END_VAR
(****************************************************************************************************)
(* CONFIGURATION: origin on the floor at the right belt edge, local +Y across the belt               *)
(****************************************************************************************************)
TempPose.fX := lr_REJECT_X;
TempPose.fY := lr_OUTFEED_Y - DEMO_GlobalConst.DEMO_lr_BELT_WIDTH / 2 - lr_GAP;
TempPose.fZ := 0;
fb_RejectUnit.m_SetPose(vi_Pose := TempPose);
TempPose.fX := 0;
TempPose.fY := -lr_HOUSING_WIDTH / 2;
TempPose.fZ := 0;
fb_RejectUnit.m_SetBody(vi_un_Body := 1, vi_e_Shape := E_VisuBodyShape.BOX, vi_e_Role := E_VisuBodyRole.STRUCTURE,
	vi_Pose := TempPose, vi_lr_Length := lr_HOUSING_LENGTH, vi_lr_Width := lr_HOUSING_WIDTH,
	vi_lr_Height := DEMO_GlobalConst.DEMO_lr_BELT_Z + lr_HOUSING_ABOVE_BELT, vi_lr_TopLength := 0, vi_lr_TopWidth := 0);
TempPose.fY := lr_PUSHER_WIDTH / 2;
TempPose.fZ := DEMO_GlobalConst.DEMO_lr_BELT_Z + lr_PUSHER_ABOVE_BELT;
fb_RejectUnit.m_SetBody(vi_un_Body := 2, vi_e_Shape := E_VisuBodyShape.BOX, vi_e_Role := E_VisuBodyRole.STRUCTURE,
	vi_Pose := TempPose, vi_lr_Length := lr_PUSHER_LENGTH, vi_lr_Width := lr_PUSHER_WIDTH, vi_lr_Height := lr_PUSHER_HEIGHT,
	vi_lr_TopLength := 0, vi_lr_TopWidth := 0);
(* The outfeed counts from its shifted origin. *)
fb_RejectUnit.m_SetZone(vi_un_Zone := 1, vi_udn_ConveyorId := fb_Outfeed.m_Id(), vi_lr_Start := lr_REJECT_X - lr_OUTFEED_ORIGIN_X,
	vi_lr_End := lr_REJECT_X - lr_OUTFEED_ORIGIN_X, vi_lr_AllocationOffset := 0,
	vi_lr_CcsOffset := lr_REJECT_X - lr_OUTFEED_ORIGIN_X, vi_lr_StartY := 0, vi_lr_EndY := 0);


(****************************************************************************************************)
(* PUSHING                                                                                          *)
(****************************************************************************************************)
IF udn_RejectPushing <> 0 THEN
	lr_RejectLeft := lr_RejectLeft - lr_Dt;
	IF lr_RejectLeft <= 0 THEN
		fb_Outfeed.m_RemoveProduct(udn_RejectPushing);
		udn_RejectPushing := 0;
	END_IF
END_IF

(* A product passes the pusher in the cycle its centre crosses lr_REJECT_X. *)
un_TempIndex := 0;
WHILE un_TempIndex < fb_Outfeed.m_ProductCount() DO
	fb_Outfeed.m_GetProduct(vi_un_Index := un_TempIndex, vo_Product => TempProduct, vo_Pose => TempProductPose);
	TempProductPose := fb_Outfeed.m_BeltToMcs(vi_Pose := TempProductPose);
	IF TempProduct.eState = E_VisuProductState.PLACED AND TempProductPose.fX >= lr_REJECT_X
		AND TempProductPose.fX - lr_OUTFEED_SPEED * lr_Dt < lr_REJECT_X
	THEN
		un_RejectPassed := un_RejectPassed + 1;
		IF un_RejectPassed MOD un_REJECT_EVERY = 0 AND udn_RejectPushing = 0 THEN
			fb_Outfeed.m_SetProductState(vi_udn_Id := TempProduct.nId, vi_e_State := E_VisuProductState.REJECTED,
				vi_udn_ClientId := fb_RejectUnit.m_Id(), vi_udn_MoverId := 0, vi_udn_FingerId := 0);
			udn_RejectPushing := TempProduct.nId;
			lr_RejectLeft := lr_REJECT_PUSH_TIME;
		END_IF
	END_IF
	un_TempIndex := un_TempIndex + 1;
END_WHILE
fb_RejectUnit.m_SetBodyActive(vi_un_Body := 2, vi_b_Active := udn_RejectPushing <> 0);
m_RejectUnit := TRUE;
END_METHOD

(****************************************************************************************************<br>
© Syntegon Group.<br>
All rights reserved, also regarding any disposal, exploitation, reproduction, editing, distribution,<br>
as well as in the event of applications for industrial property rights.<br>
*****************************************************************************************************<br>
DESCRIPTION:<br>
Moves the Delta 3 fingers and reports the TCP, the fault and the finger states of Delta n_Robot.<br>
****************************************************************************************************)
METHOD PRIVATE m_Report : BOOL
(* Delta 3 closes its fingers while it descends onto a product and keeps them closed while it carries one. *)
IF n_Robot = 2 THEN
	IF n_Phase[n_Robot] = n_PHASE_DESCEND OR n_HeldCount[n_Robot] > 0 THEN
		lr_Spread := _FC_DemoApproach(lr_Spread, lr_SpreadClosed, lr_SPREAD_SPEED * lr_Dt);
	ELSE
		lr_Spread := _FC_DemoApproach(lr_Spread, lr_SPREAD_OPEN, lr_SPREAD_SPEED * lr_Dt);
	END_IF
END_IF

(* Only the TCP (the flange) is reported; the visualisation derives the arms. A small offset shows the setpoint
   marker. Tool rotations show only through the finger poses. *)
SetpointTcp := Tcp[n_Robot];
SetpointTcp.fX := SetpointTcp.fX + 2;
SetpointTcp.fZ := SetpointTcp.fZ - 1;
fb_RefRobot.m_SetTcp(vi_ActualTcp := Tcp[n_Robot], vi_SetpointTcp := SetpointTcp);

(* Demo fault: Delta 1 overheats now and then; a Reset acknowledges it until the next fault period. *)
IF n_Robot = 0 AND DEMO_GlobalVar.DEMO_lr_FaultPhase < lr_FAULT_START THEN
	b_FaultAcknowledged := FALSE;
END_IF
fb_RefRobot.m_SetFault(vi_b_Active := n_Robot = 0 AND NOT b_FaultAcknowledged AND DEMO_GlobalVar.DEMO_lr_FaultPhase >= lr_FAULT_START
										AND DEMO_GlobalVar.DEMO_lr_FaultPhase
											< lr_FAULT_START + DEMO_GlobalConst.DEMO_lr_FAULT_DURATION,
	vi_str_Message := 'Drive 2: overtemperature');
FOR n_Finger := 1 TO n_FingerCount DO
	(* Delta 1: a cup grips while its slot holds a product; the others grip while anything is carried. *)
	fb_RefRobot.m_SetFingerState(vi_un_Finger := INT_TO_UINT(n_Finger),
		vi_Pose := m_FingerPose(vi_n_Robot := n_Robot, vi_n_Finger := n_Finger),
		vi_b_Active := n_HeldCount[n_Robot] >= SEL(n_Robot = 0, 1, n_Finger));
END_FOR
m_Report := TRUE;
END_METHOD

(****************************************************************************************************<br>
© Syntegon Group.<br>
All rights reserved, also regarding any disposal, exploitation, reproduction, editing, distribution,<br>
as well as in the event of applications for industrial property rights.<br>
*****************************************************************************************************<br>
DESCRIPTION:<br>
Reset of the machine (accepted while stopped): every product leaves Infeed 1's register, no robot approaches or<br>
carries one of its products any more (Delta 1 nothing at all), the generator starts again from its seed, the<br>
missed-product message and Delta 1's fault are acknowledged.<br>
****************************************************************************************************)
METHOD PRIVATE m_Reset : BOOL
VAR
	n_TempRobot							: INT;
	n_TempSlot							: INT;
	b_TempFromInfeed1					: BOOL;	// [-] the robot carries a product of Infeed 1
	TempProduct							: ST_VisuProduct;
	TempPose							: ST_VisuPlanarPose;
END_VAR
WHILE fb_Infeed1.m_ProductCount() > 0 DO
	fb_Infeed1.m_GetProduct(vi_un_Index := 0, vo_Product => TempProduct, vo_Pose => TempPose);
	IF NOT fb_Infeed1.m_RemoveProduct(TempProduct.nId) THEN
		EXIT;	// never: the first entry is always there
	END_IF
END_WHILE
FOR n_TempRobot := 0 TO 2 DO
	b_TempFromInfeed1 := FALSE;
	FOR n_TempSlot := 0 TO n_HeldCount[n_TempRobot] - 1 DO
		b_TempFromInfeed1 := b_TempFromInfeed1 OR n_HeldBelt[n_TempRobot, n_TempSlot] = 0;
	END_FOR
	IF n_TempRobot = 0 OR b_TempFromInfeed1 OR (udn_TargetId[n_TempRobot] <> 0 AND n_TargetBelt[n_TempRobot] = 0) THEN
		udn_TargetId[n_TempRobot] := 0;
		n_HeldCount[n_TempRobot] := 0;
		n_Phase[n_TempRobot] := n_PHASE_IDLE;
	END_IF
END_FOR
dn_GenSeed := 0;	// the generator starts again from the recipe's seed
lr_MissedLeft := 0;
b_FaultAcknowledged := TRUE;
m_Reset := TRUE;
END_METHOD

(****************************************************************************************************<br>
© Syntegon Group.<br>
All rights reserved, also regarding any disposal, exploitation, reproduction, editing, distribution,<br>
as well as in the event of applications for industrial property rights.<br>
*****************************************************************************************************<br>
DESCRIPTION:<br>
Pick and place sequence of Delta n_Robot: allocate, approach, descend and pick, lift (Delta 1 picks twice),<br>
transfer to the outfeed, lower and release every carried product.<br>
****************************************************************************************************)
METHOD PRIVATE m_Sequence : BOOL
CASE n_Phase[n_Robot] OF
	n_PHASE_IDLE:
		IF NOT m_Allocate() THEN
			m_MoveToward(vio_Tcp := Tcp[n_Robot], vi_lr_TargetX := lr_BaseX, vi_lr_TargetY := lr_ROBOT_Y,
				vi_lr_TargetZ := lr_ROBOT_Z - 900, vi_lr_MaxStep := lr_Step);
		END_IF

	n_PHASE_APPROACH:
		IF lr_X - lr_LEAD > lr_BaseX + lr_PICK_HALF_ZONE THEN
			(* Product left the zone: hand it back, a downstream robot may still catch it. *)
			fb_RefBelt.m_SetProductState(vi_udn_Id := udn_TargetId[n_Robot], vi_e_State := E_VisuProductState.DETECTED,
				vi_udn_ClientId := fb_RefRobot.m_Id(), vi_udn_MoverId := 0, vi_udn_FingerId := 0);
			udn_TargetId[n_Robot] := 0;
			n_Phase[n_Robot] := n_PHASE_IDLE;
		ELSE
			lr_ToolRz[n_Robot] := lr_ToolRz[n_Robot] + (lr_TargetRz - lr_ToolRz[n_Robot]) * MIN(1.0, lr_Dt * 10.0);
			IF m_MoveToward(vio_Tcp := Tcp[n_Robot], vi_lr_TargetX := lr_X - Grip.fX, vi_lr_TargetY := lr_Y - Grip.fY,
				vi_lr_TargetZ := lr_TopZ - Grip.fZ + lr_HOVER, vi_lr_MaxStep := lr_Step)
			THEN
				n_Phase[n_Robot] := n_PHASE_DESCEND;
			END_IF
		END_IF

	n_PHASE_DESCEND:
		lr_ToolRz[n_Robot] := lr_ToolRz[n_Robot] + (lr_TargetRz - lr_ToolRz[n_Robot]) * MIN(1.0, lr_Dt * 10.0);
		(* Delta 3 grips only once its fingers have closed around the product (both operands are evaluated). *)
		IF m_MoveToward(vio_Tcp := Tcp[n_Robot], vi_lr_TargetX := lr_X - Grip.fX, vi_lr_TargetY := lr_Y - Grip.fY,
			vi_lr_TargetZ := lr_TopZ - Grip.fZ, vi_lr_MaxStep := lr_Step)
		AND (n_Robot <> 2 OR lr_Spread = lr_SpreadClosed)
		THEN
			n_Slot := n_HeldCount[n_Robot];
			fb_RefBelt.m_SetProductState(vi_udn_Id := udn_TargetId[n_Robot], vi_e_State := E_VisuProductState.PICKED,
				vi_udn_ClientId := fb_RefRobot.m_Id(), vi_udn_MoverId := 0, vi_udn_FingerId := INT_TO_UDINT(n_Finger));
			udn_Held[n_Robot, n_Slot] := udn_TargetId[n_Robot];
			n_HeldBelt[n_Robot, n_Slot] := n_TargetBelt[n_Robot];
			udn_HeldType[n_Robot, n_Slot] := Product.nProductType;
			un_HeldMark[n_Robot, n_Slot] := Product.nMark;
			n_HeldCount[n_Robot] := n_Slot + 1;
			udn_TargetId[n_Robot] := 0;
			n_Phase[n_Robot] := n_PHASE_LIFT;
		END_IF

	n_PHASE_LIFT:
		IF m_MoveToward(vio_Tcp := Tcp[n_Robot], vi_lr_TargetX := Tcp[n_Robot].fX, vi_lr_TargetY := Tcp[n_Robot].fY,
			vi_lr_TargetZ := DEMO_GlobalConst.DEMO_lr_BELT_Z + lr_HeldHeight + lr_GripHeight
							+ lr_HOVER,
			vi_lr_MaxStep := lr_Step)
		THEN
			(* Delta 1 picks as many products as its recipe says (1 or 2, one per cup) before it places them. *)
			IF n_Robot = 0 AND n_HeldCount[n_Robot] < LIMIT(1, DEMO_GlobalVar.DEMO_Recipe.dn_PicksPerCycle, 2) THEN
				n_Phase[n_Robot] := n_PHASE_IDLE;
			ELSE
				n_Phase[n_Robot] := n_PHASE_TRANSFER;
			END_IF
		END_IF

	n_PHASE_TRANSFER:
		lr_ToolRz[n_Robot] := lr_ToolRz[n_Robot] * (1.0 - MIN(1.0, lr_Dt * 5.0));
		IF n_Robot = 1 THEN
			lr_TiltRx := _FC_DemoApproach(lr_TiltRx, lr_TILT_ANGLE, lr_TILT_SPEED * lr_Dt);
		END_IF
		(* Now and then Delta 2 places far downstream and waits there for a gap on the outfeed: a real limit
		   violation for the visualisation, its TCP limit area in Delta 3's limit area meanwhile. *)
		b_FarPlace := n_Robot = 1 AND un_Placed[n_Robot] MOD un_FAR_PLACE_EVERY = un_FAR_PLACE_EVERY - 1;
		IF m_MoveToward(vio_Tcp := Tcp[n_Robot], vi_lr_TargetX := lr_BaseX + SEL(b_FarPlace, 0, lr_FAR_PLACE_OFFSET),
			vi_lr_TargetY := lr_OUTFEED_Y,
			vi_lr_TargetZ := DEMO_GlobalConst.DEMO_lr_BELT_Z + lr_HeldHeight + lr_GripHeight
							+ lr_HOVER,
			vi_lr_MaxStep := lr_Step)
		THEN
			lr_PlaceWait[n_Robot] := lr_PlaceWait[n_Robot] + lr_Dt;
			IF NOT b_FarPlace OR lr_PlaceWait[n_Robot] >= lr_FAR_PLACE_WAIT THEN
				lr_PlaceWait[n_Robot] := 0;
				n_Phase[n_Robot] := n_PHASE_LOWER;
			END_IF
		END_IF

